(* IEC 61131-3 sources: plc-st-coding-agent/progress/evidence/f14_v3_parallel_20261112/jobs/codex_minimax-m27, 122 files *)

(* ---- public-easy-01.candidate_01.st ---- *)
FUNCTION_BLOCK FillingLineControl
VAR
    currentState : INT := 0;
END_VAR

CASE currentState OF
    0:
        Pump_Motor := FALSE;
        Filling_Valve := FALSE;
        Capping_Machine := FALSE;
        Packing_Machine := FALSE;
        Completion_Light := FALSE;

        IF bottleSensor THEN
            currentState := 1;
        END_IF;

    1:
        Pump_Motor := TRUE;

        IF cleaningConfirmButton THEN
            currentState := 2;
        END_IF;

    2:
        Pump_Motor := FALSE;
        Filling_Valve := TRUE;

        IF fillingConfirmButton THEN
            currentState := 3;
        END_IF;

    3:
        Filling_Valve := FALSE;
        Capping_Machine := TRUE;

        IF cappingConfirmButton THEN
            currentState := 4;
        END_IF;

    4:
        Capping_Machine := FALSE;
        Packing_Machine := TRUE;

        IF packingConfirmButton THEN
            currentState := 5;
        END_IF;

    5:
        Packing_Machine := FALSE;
        Completion_Light := TRUE;

        IF finishedButton THEN
            currentState := 0;
        END_IF;
END_CASE;
END_FUNCTION_BLOCK

(* ---- public-easy-01.candidate_02.st ---- *)
FUNCTION_BLOCK FillingLineControl
VAR_INPUT
    bottleSensor : BOOL;
    cleaningConfirmButton : BOOL;
    fillingConfirmButton : BOOL;
    cappingConfirmButton : BOOL;
    packingConfirmButton : BOOL;
    finishedButton : BOOL;
END_VAR
VAR_OUTPUT
    Pump_Motor : BOOL;
    Filling_Valve : BOOL;
    Capping_Machine : BOOL;
    Packing_Machine : BOOL;
    Completion_Light : BOOL;
END_VAR
VAR
    currentState : INT := 0;
END_VAR

CASE currentState OF
    0:
        Pump_Motor := FALSE;
        Filling_Valve := FALSE;
        Capping_Machine := FALSE;
        Packing_Machine := FALSE;
        Completion_Light := FALSE;

        IF bottleSensor THEN
            currentState := 1;
        END_IF;

    1:
        Pump_Motor := TRUE;

        IF cleaningConfirmButton THEN
            currentState := 2;
        END_IF;

    2:
        Pump_Motor := FALSE;
        Filling_Valve := TRUE;

        IF fillingConfirmButton THEN
            currentState := 3;
        END_IF;

    3:
        Filling_Valve := FALSE;
        Capping_Machine := TRUE;

        IF cappingConfirmButton THEN
            currentState := 4;
        END_IF;

    4:
        Capping_Machine := FALSE;
        Packing_Machine := TRUE;

        IF packingConfirmButton THEN
            currentState := 5;
        END_IF;

    5:
        Packing_Machine := FALSE;
        Completion_Light := TRUE;

        IF finishedButton THEN
            currentState := 0;
        END_IF;
END_CASE;
END_FUNCTION_BLOCK

(* ---- public-easy-01.raw_candidate_01.st ---- *)
FUNCTION_BLOCK FillingLineControl
VAR
    currentState : INT := 0;
END_VAR

CASE currentState OF
    0:
        Pump_Motor := FALSE;
        Filling_Valve := FALSE;
        Capping_Machine := FALSE;
        Packing_Machine := FALSE;
        Completion_Light := FALSE;

        IF bottleSensor THEN
            currentState := 1;
        END_IF;

    1:
        Pump_Motor := TRUE;

        IF cleaningConfirmButton THEN
            currentState := 2;
        END_IF;

    2:
        Pump_Motor := FALSE;
        Filling_Valve := TRUE;

        IF fillingConfirmButton THEN
            currentState := 3;
        END_IF;

    3:
        Filling_Valve := FALSE;
        Capping_Machine := TRUE;

        IF cappingConfirmButton THEN
            currentState := 4;
        END_IF;

    4:
        Capping_Machine := FALSE;
        Packing_Machine := TRUE;

        IF packingConfirmButton THEN
            currentState := 5;
        END_IF;

    5:
        Packing_Machine := FALSE;
        Completion_Light := TRUE;

        IF finishedButton THEN
            currentState := 0;
        END_IF;
END_CASE;
END_FUNCTION_BLOCK

(* ---- public-easy-01.raw_candidate_02.st ---- *)
FUNCTION_BLOCK FillingLineControl
VAR_INPUT
    bottleSensor : BOOL;
    cleaningConfirmButton : BOOL;
    fillingConfirmButton : BOOL;
    cappingConfirmButton : BOOL;
    packingConfirmButton : BOOL;
    finishedButton : BOOL;
END_VAR
VAR_OUTPUT
    Pump_Motor : BOOL;
    Filling_Valve : BOOL;
    Capping_Machine : BOOL;
    Packing_Machine : BOOL;
    Completion_Light : BOOL;
END_VAR
VAR
    currentState : INT := 0;
END_VAR

CASE currentState OF
    0:
        Pump_Motor := FALSE;
        Filling_Valve := FALSE;
        Capping_Machine := FALSE;
        Packing_Machine := FALSE;
        Completion_Light := FALSE;

        IF bottleSensor THEN
            currentState := 1;
        END_IF;

    1:
        Pump_Motor := TRUE;

        IF cleaningConfirmButton THEN
            currentState := 2;
        END_IF;

    2:
        Pump_Motor := FALSE;
        Filling_Valve := TRUE;

        IF fillingConfirmButton THEN
            currentState := 3;
        END_IF;

    3:
        Filling_Valve := FALSE;
        Capping_Machine := TRUE;

        IF cappingConfirmButton THEN
            currentState := 4;
        END_IF;

    4:
        Capping_Machine := FALSE;
        Packing_Machine := TRUE;

        IF packingConfirmButton THEN
            currentState := 5;
        END_IF;

    5:
        Packing_Machine := FALSE;
        Completion_Light := TRUE;

        IF finishedButton THEN
            currentState := 0;
        END_IF;
END_CASE;
END_FUNCTION_BLOCK

(* ---- public-easy-02.candidate_01.st ---- *)
FUNCTION_BLOCK FB_DualWordEdgeDetection
VAR_INPUT
END_VAR

VAR_OUTPUT
    hasChanged       : BOOL  := FALSE;
    hasRisingEdges   : BOOL  := FALSE;
    risingBits       : DWORD := 0;
    noOfRisingBits   : USINT := 0;
    hasFallingEdges  : BOOL  := FALSE;
    fallingBits      : DWORD := 0;
    noOfFallingBits  : USINT := 0;
END_VAR

VAR
    prevValue : DWORD := 0;
    bitMask   : DWORD;
    bitCount  : USINT;
END_VAR

// Detect rising edges: current=1 AND previous=0
risingBits := value AND (NOT prevValue);

// Detect falling edges: current=0 AND previous=1
fallingBits := (NOT value) AND prevValue;

// Set change indicators
hasChanged := (risingBits OR fallingBits) <> 0;
hasRisingEdges := risingBits <> 0;
hasFallingEdges := fallingBits <> 0;

// Count rising bits
bitMask := risingBits;
noOfRisingBits := 0;
FOR bitCount := 0 TO 31 DO
    IF (bitMask AND 1) = 1 THEN
        noOfRisingBits := noOfRisingBits + 1;
    END_IF;
    bitMask := SHR(bitMask, 1);
END_FOR;

// Count falling bits
bitMask := fallingBits;
noOfFallingBits := 0;
FOR bitCount := 0 TO 31 DO
    IF (bitMask AND 1) = 1 THEN
        noOfFallingBits := noOfFallingBits + 1;
    END_IF;
    bitMask := SHR(bitMask, 1);
END_FOR;

// Store current value for next scan
prevValue := value;

END_FUNCTION_BLOCK

(* ---- public-easy-02.candidate_02.st ---- *)
FUNCTION_BLOCK FB_DualWordEdgeDetection
VAR_INPUT
    value : DWORD;
END_VAR

VAR_OUTPUT
    hasChanged       : BOOL  := FALSE;
    hasRisingEdges   : BOOL  := FALSE;
    risingBits       : DWORD := 0;
    noOfRisingBits   : USINT := 0;
    hasFallingEdges  : BOOL  := FALSE;
    fallingBits      : DWORD := 0;
    noOfFallingBits  : USINT := 0;
END_VAR

VAR
    prevValue : DWORD := 0;
    tmpBits   : DWORD;
END_VAR

risingBits := value AND (NOT prevValue);
fallingBits := (NOT value) AND prevValue;

hasChanged := risingBits <> 0 OR fallingBits <> 0;
hasRisingEdges := risingBits <> 0;
hasFallingEdges := fallingBits <> 0;

tmpBits := risingBits;
noOfRisingBits := 0;
WHILE tmpBits <> 0 DO
    noOfRisingBits := noOfRisingBits + 1;
    tmpBits := SHR(tmpBits, 1);
END_WHILE;

tmpBits := fallingBits;
noOfFallingBits := 0;
WHILE tmpBits <> 0 DO
    noOfFallingBits := noOfFallingBits + 1;
    tmpBits := SHR(tmpBits, 1);
END_WHILE;

prevValue := value;

END_FUNCTION_BLOCK

(* ---- public-easy-02.raw_candidate_01.st ---- *)
FUNCTION_BLOCK FB_DualWordEdgeDetection
VAR_INPUT
END_VAR

VAR_OUTPUT
    hasChanged       : BOOL  := FALSE;
    hasRisingEdges   : BOOL  := FALSE;
    risingBits       : DWORD := 0;
    noOfRisingBits   : USINT := 0;
    hasFallingEdges  : BOOL  := FALSE;
    fallingBits      : DWORD := 0;
    noOfFallingBits  : USINT := 0;
END_VAR

VAR
    prevValue : DWORD := 0;
    bitMask   : DWORD;
    bitCount  : USINT;
END_VAR

// Detect rising edges: current=1 AND previous=0
risingBits := value AND (NOT prevValue);

// Detect falling edges: current=0 AND previous=1
fallingBits := (NOT value) AND prevValue;

// Set change indicators
hasChanged := (risingBits OR fallingBits) <> 0;
hasRisingEdges := risingBits <> 0;
hasFallingEdges := fallingBits <> 0;

// Count rising bits
bitMask := risingBits;
noOfRisingBits := 0;
FOR bitCount := 0 TO 31 DO
    IF (bitMask AND 1) = 1 THEN
        noOfRisingBits := noOfRisingBits + 1;
    END_IF;
    bitMask := SHR(bitMask, 1);
END_FOR;

// Count falling bits
bitMask := fallingBits;
noOfFallingBits := 0;
FOR bitCount := 0 TO 31 DO
    IF (bitMask AND 1) = 1 THEN
        noOfFallingBits := noOfFallingBits + 1;
    END_IF;
    bitMask := SHR(bitMask, 1);
END_FOR;

// Store current value for next scan
prevValue := value;

END_FUNCTION_BLOCK

(* ---- public-easy-02.raw_candidate_02.st ---- *)
FUNCTION_BLOCK FB_DualWordEdgeDetection
VAR_INPUT
    value : DWORD;
END_VAR

VAR_OUTPUT
    hasChanged       : BOOL  := FALSE;
    hasRisingEdges   : BOOL  := FALSE;
    risingBits       : DWORD := 0;
    noOfRisingBits   : USINT := 0;
    hasFallingEdges  : BOOL  := FALSE;
    fallingBits      : DWORD := 0;
    noOfFallingBits  : USINT := 0;
END_VAR

VAR
    prevValue : DWORD := 0;
    tmpBits   : DWORD;
END_VAR

risingBits := value AND (NOT prevValue);
fallingBits := (NOT value) AND prevValue;

hasChanged := risingBits <> 0 OR fallingBits <> 0;
hasRisingEdges := risingBits <> 0;
hasFallingEdges := fallingBits <> 0;

tmpBits := risingBits;
noOfRisingBits := 0;
WHILE tmpBits <> 0 DO
    noOfRisingBits := noOfRisingBits + 1;
    tmpBits := SHR(tmpBits, 1);
END_WHILE;

tmpBits := fallingBits;
noOfFallingBits := 0;
WHILE tmpBits <> 0 DO
    noOfFallingBits := noOfFallingBits + 1;
    tmpBits := SHR(tmpBits, 1);
END_WHILE;

prevValue := value;

END_FUNCTION_BLOCK

(* ---- public-easy-04.candidate_01.st ---- *)
FUNCTION_BLOCK JamPumpControl
VAR_INPUT
    VISCOSITY_OK     : BOOL;
    PASTE_E_STOP_NC  : BOOL;
    DebounceTime     : TIME;
    CycleTime        : TIME;
END_VAR

VAR_OUTPUT
    VFD_RUN          : BOOL := FALSE;
    PUMP_MAINT_DUE   : BOOL := FALSE;
    PUMP_RUNTIME_ACC : LTIME := LTIME#0s;
END_VAR

VAR
    ViscosityValid        : BOOL := FALSE;
    ViscosityDebounceTmr  : LTIME := LTIME#0s;
END_VAR

// Viscosity debouncing
IF VISCOSITY_OK THEN
    IF NOT ViscosityValid THEN
        ViscosityDebounceTmr := ViscosityDebounceTmr + LTIME(CycleTime);
        IF ViscosityDebounceTmr >= LTIME(DebounceTime) THEN
            ViscosityValid := TRUE;
            ViscosityDebounceTmr := LTIME#0s;
        END_IF;
    END_IF;
ELSE
    ViscosityValid := FALSE;
    ViscosityDebounceTmr := LTIME#0s;
END_IF;

// Safety permissive: E-stop AND valid viscosity
IF PASTE_E_STOP_NC AND ViscosityValid THEN
    VFD_RUN := TRUE;
ELSE
    VFD_RUN := FALSE;
END_IF;

// Runtime accumulation while running
IF VFD_RUN THEN
    PUMP_RUNTIME_ACC := PUMP_RUNTIME_ACC + LTIME(CycleTime);
END_IF;

// Maintenance due at 500 hours
PUMP_MAINT_DUE := (PUMP_RUNTIME_ACC >= LTIME#500h);

END_FUNCTION_BLOCK

(* ---- public-easy-04.candidate_02.st ---- *)
FUNCTION_BLOCK JamPumpControl
VAR_INPUT
    VISCOSITY_OK    : BOOL;
    PASTE_E_STOP_NC : BOOL;
    DebounceTime    : TIME;
    CycleTime       : TIME;
END_VAR

VAR_OUTPUT
    VFD_RUN          : BOOL := FALSE;
    PUMP_MAINT_DUE   : BOOL := FALSE;
    PUMP_RUNTIME_ACC : LTIME := LTIME#0s;
END_VAR

VAR
    ViscosityValid       : BOOL := FALSE;
    ViscosityDebounceTmr : LTIME := LTIME#0s;
END_VAR

IF VISCOSITY_OK THEN
    IF NOT ViscosityValid THEN
        ViscosityDebounceTmr := ViscosityDebounceTmr + CycleTime;
        IF ViscosityDebounceTmr >= DebounceTime THEN
            ViscosityValid := TRUE;
            ViscosityDebounceTmr := LTIME#0s;
        END_IF;
    END_IF;
ELSE
    ViscosityValid := FALSE;
    ViscosityDebounceTmr := LTIME#0s;
END_IF;

IF PASTE_E_STOP_NC AND ViscosityValid THEN
    VFD_RUN := TRUE;
ELSE
    VFD_RUN := FALSE;
END_IF;

IF VFD_RUN THEN
    PUMP_RUNTIME_ACC := PUMP_RUNTIME_ACC + CycleTime;
END_IF;

PUMP_MAINT_DUE := (PUMP_RUNTIME_ACC >= LTIME#500h);

END_FUNCTION_BLOCK

(* ---- public-easy-04.raw_candidate_01.st ---- *)
FUNCTION_BLOCK JamPumpControl
VAR_INPUT
    VISCOSITY_OK     : BOOL;
    PASTE_E_STOP_NC  : BOOL;
    DebounceTime     : TIME;
    CycleTime        : TIME;
END_VAR

VAR_OUTPUT
    VFD_RUN          : BOOL := FALSE;
    PUMP_MAINT_DUE   : BOOL := FALSE;
    PUMP_RUNTIME_ACC : LTIME := LTIME#0s;
END_VAR

VAR
    ViscosityValid        : BOOL := FALSE;
    ViscosityDebounceTmr  : LTIME := LTIME#0s;
END_VAR

// Viscosity debouncing
IF VISCOSITY_OK THEN
    IF NOT ViscosityValid THEN
        ViscosityDebounceTmr := ViscosityDebounceTmr + LTIME(CycleTime);
        IF ViscosityDebounceTmr >= LTIME(DebounceTime) THEN
            ViscosityValid := TRUE;
            ViscosityDebounceTmr := LTIME#0s;
        END_IF;
    END_IF;
ELSE
    ViscosityValid := FALSE;
    ViscosityDebounceTmr := LTIME#0s;
END_IF;

// Safety permissive: E-stop AND valid viscosity
IF PASTE_E_STOP_NC AND ViscosityValid THEN
    VFD_RUN := TRUE;
ELSE
    VFD_RUN := FALSE;
END_IF;

// Runtime accumulation while running
IF VFD_RUN THEN
    PUMP_RUNTIME_ACC := PUMP_RUNTIME_ACC + LTIME(CycleTime);
END_IF;

// Maintenance due at 500 hours
PUMP_MAINT_DUE := (PUMP_RUNTIME_ACC >= LTIME#500h);

END_FUNCTION_BLOCK

(* ---- public-easy-04.raw_candidate_02.st ---- *)
FUNCTION_BLOCK JamPumpControl
VAR_INPUT
    VISCOSITY_OK    : BOOL;
    PASTE_E_STOP_NC : BOOL;
    DebounceTime    : TIME;
    CycleTime       : TIME;
END_VAR

VAR_OUTPUT
    VFD_RUN          : BOOL := FALSE;
    PUMP_MAINT_DUE   : BOOL := FALSE;
    PUMP_RUNTIME_ACC : LTIME := LTIME#0s;
END_VAR

VAR
    ViscosityValid       : BOOL := FALSE;
    ViscosityDebounceTmr : LTIME := LTIME#0s;
END_VAR

IF VISCOSITY_OK THEN
    IF NOT ViscosityValid THEN
        ViscosityDebounceTmr := ViscosityDebounceTmr + CycleTime;
        IF ViscosityDebounceTmr >= DebounceTime THEN
            ViscosityValid := TRUE;
            ViscosityDebounceTmr := LTIME#0s;
        END_IF;
    END_IF;
ELSE
    ViscosityValid := FALSE;
    ViscosityDebounceTmr := LTIME#0s;
END_IF;

IF PASTE_E_STOP_NC AND ViscosityValid THEN
    VFD_RUN := TRUE;
ELSE
    VFD_RUN := FALSE;
END_IF;

IF VFD_RUN THEN
    PUMP_RUNTIME_ACC := PUMP_RUNTIME_ACC + CycleTime;
END_IF;

PUMP_MAINT_DUE := (PUMP_RUNTIME_ACC >= LTIME#500h);

END_FUNCTION_BLOCK

(* ---- public-easy-05.candidate_01.st ---- *)
FUNCTION_BLOCK WeldGapAlarm
VAR_INPUT
    Gap_Exceeded : BOOL;
    Weld_E_Stop_NC : BOOL;
    DebounceTime : TIME;
END_VAR

VAR_OUTPUT
    Operator_Alert : BOOL := FALSE;
    Weld_Soft_Start_Active : BOOL := TRUE;
END_VAR

VAR
    initTimer : TON;
    debounceTimer : TON;
    monitoringActive : BOOL := FALSE;
END_VAR

// E-Stop takes priority over all states
IF NOT Weld_E_Stop_NC THEN
    Operator_Alert := FALSE;
    Weld_Soft_Start_Active := FALSE;
    monitoringActive := FALSE;

    // Reset timers when E-Stop is active
    initTimer(IN := FALSE);
    debounceTimer(IN := FALSE);
    initTimer();
    debounceTimer();
    RETURN;
END_IF;

// Initialization phase: 5-second power-up inhibition
IF NOT monitoringActive THEN
    initTimer(IN := TRUE, PT := T#5S);
    initTimer();

    Operator_Alert := FALSE;
    Weld_Soft_Start_Active := TRUE;

    IF initTimer.Q THEN
        monitoringActive := TRUE;
        Weld_Soft_Start_Active := FALSE;

        // Reset timers upon entering monitoring
        initTimer(IN := FALSE);
        debounceTimer(IN := FALSE);
        initTimer();
        debounceTimer();
    END_IF;

    initTimer(IN := FALSE);
    initTimer();
    RETURN;
END_IF;

// Normal gap monitoring with debounce
IF NOT Gap_Exceeded THEN
    Operator_Alert := FALSE;
    debounceTimer(IN := FALSE);
    debounceTimer();
ELSE
    debounceTimer(IN := TRUE, PT := DebounceTime);
    debounceTimer();

    IF debounceTimer.Q THEN
        Operator_Alert := TRUE;
    END_IF;
END_IF;

END_FUNCTION_BLOCK

(* ---- public-easy-05.candidate_02.st ---- *)
FUNCTION_BLOCK WeldGapAlarm
VAR_INPUT
    Gap_Exceeded : BOOL;
    Weld_E_Stop_NC : BOOL;
    DebounceTime : TIME;
END_VAR

VAR_OUTPUT
    Operator_Alert : BOOL := FALSE;
    Weld_Soft_Start_Active : BOOL := TRUE;
END_VAR

VAR
    initTimer : TON;
    debounceTimer : TON;
    state : UINT := 0;
END_VAR

IF NOT Weld_E_Stop_NC THEN
    Operator_Alert := FALSE;
    Weld_Soft_Start_Active := FALSE;
    state := 0;
    initTimer(IN := FALSE);
    debounceTimer(IN := FALSE);
    initTimer();
    debounceTimer();
    RETURN;
END_IF;

IF state = 0 THEN
    initTimer(IN := TRUE, PT := T#5S);
    initTimer();
    Operator_Alert := FALSE;
    Weld_Soft_Start_Active := TRUE;

    IF initTimer.Q THEN
        state := 1;
        initTimer(IN := FALSE);
        debounceTimer(IN := FALSE);
        initTimer();
        debounceTimer();
    END_IF;
    RETURN;
END_IF;

IF state = 1 THEN
    Weld_Soft_Start_Active := FALSE;

    IF NOT Gap_Exceeded THEN
        Operator_Alert := FALSE;
        debounceTimer(IN := FALSE);
        debounceTimer();
    ELSE
        debounceTimer(IN := TRUE, PT := DebounceTime);
        debounceTimer();

        IF debounceTimer.Q THEN
            Operator_Alert := TRUE;
        END_IF;
    END_IF;
END_IF;

END_FUNCTION_BLOCK

(* ---- public-easy-05.raw_candidate_01.st ---- *)
FUNCTION_BLOCK WeldGapAlarm
VAR_INPUT
    Gap_Exceeded : BOOL;
    Weld_E_Stop_NC : BOOL;
    DebounceTime : TIME;
END_VAR

VAR_OUTPUT
    Operator_Alert : BOOL := FALSE;
    Weld_Soft_Start_Active : BOOL := TRUE;
END_VAR

VAR
    initTimer : TON;
    debounceTimer : TON;
    monitoringActive : BOOL := FALSE;
END_VAR

// E-Stop takes priority over all states
IF NOT Weld_E_Stop_NC THEN
    Operator_Alert := FALSE;
    Weld_Soft_Start_Active := FALSE;
    monitoringActive := FALSE;

    // Reset timers when E-Stop is active
    initTimer(IN := FALSE);
    debounceTimer(IN := FALSE);
    initTimer();
    debounceTimer();
    RETURN;
END_IF;

// Initialization phase: 5-second power-up inhibition
IF NOT monitoringActive THEN
    initTimer(IN := TRUE, PT := T#5S);
    initTimer();

    Operator_Alert := FALSE;
    Weld_Soft_Start_Active := TRUE;

    IF initTimer.Q THEN
        monitoringActive := TRUE;
        Weld_Soft_Start_Active := FALSE;

        // Reset timers upon entering monitoring
        initTimer(IN := FALSE);
        debounceTimer(IN := FALSE);
        initTimer();
        debounceTimer();
    END_IF;

    initTimer(IN := FALSE);
    initTimer();
    RETURN;
END_IF;

// Normal gap monitoring with debounce
IF NOT Gap_Exceeded THEN
    Operator_Alert := FALSE;
    debounceTimer(IN := FALSE);
    debounceTimer();
ELSE
    debounceTimer(IN := TRUE, PT := DebounceTime);
    debounceTimer();

    IF debounceTimer.Q THEN
        Operator_Alert := TRUE;
    END_IF;
END_IF;

END_FUNCTION_BLOCK

(* ---- public-easy-05.raw_candidate_02.st ---- *)
FUNCTION_BLOCK WeldGapAlarm
VAR_INPUT
    Gap_Exceeded : BOOL;
    Weld_E_Stop_NC : BOOL;
    DebounceTime : TIME;
END_VAR

VAR_OUTPUT
    Operator_Alert : BOOL := FALSE;
    Weld_Soft_Start_Active : BOOL := TRUE;
END_VAR

VAR
    initTimer : TON;
    debounceTimer : TON;
    state : UINT := 0;
END_VAR

IF NOT Weld_E_Stop_NC THEN
    Operator_Alert := FALSE;
    Weld_Soft_Start_Active := FALSE;
    state := 0;
    initTimer(IN := FALSE);
    debounceTimer(IN := FALSE);
    initTimer();
    debounceTimer();
    RETURN;
END_IF;

IF state = 0 THEN
    initTimer(IN := TRUE, PT := T#5S);
    initTimer();
    Operator_Alert := FALSE;
    Weld_Soft_Start_Active := TRUE;

    IF initTimer.Q THEN
        state := 1;
        initTimer(IN := FALSE);
        debounceTimer(IN := FALSE);
        initTimer();
        debounceTimer();
    END_IF;
    RETURN;
END_IF;

IF state = 1 THEN
    Weld_Soft_Start_Active := FALSE;

    IF NOT Gap_Exceeded THEN
        Operator_Alert := FALSE;
        debounceTimer(IN := FALSE);
        debounceTimer();
    ELSE
        debounceTimer(IN := TRUE, PT := DebounceTime);
        debounceTimer();

        IF debounceTimer.Q THEN
            Operator_Alert := TRUE;
        END_IF;
    END_IF;
END_IF;

END_FUNCTION_BLOCK

(* ---- public-easy-06.candidate_01.st ---- *)
FUNCTION_BLOCK AerationBlowerControl
VAR_INPUT
    DO_LOW : BOOL;
    AERATION_E_STOP_NC : BOOL;
END_VAR

VAR_OUTPUT
    BLOWER_RUN : BOOL := FALSE;
    AERATION_BLOWER_CYCLE_COUNT : UINT := 0;
END_VAR

VAR
    StartTimer : TON;
    WasRunning : BOOL := FALSE;
END_VAR

    StartTimer(IN := DO_LOW AND AERATION_E_STOP_NC, PT := T#5S);

    BLOWER_RUN := StartTimer.Q;

    IF BLOWER_RUN AND NOT WasRunning THEN
        AERATION_BLOWER_CYCLE_COUNT := AERATION_BLOWER_CYCLE_COUNT + 1;
    END_IF;

    WasRunning := BLOWER_RUN;
END_FUNCTION_BLOCK

(* ---- public-easy-06.raw_candidate_01.st ---- *)
FUNCTION_BLOCK AerationBlowerControl
VAR_INPUT
    DO_LOW : BOOL;
    AERATION_E_STOP_NC : BOOL;
END_VAR

VAR_OUTPUT
    BLOWER_RUN : BOOL := FALSE;
    AERATION_BLOWER_CYCLE_COUNT : UINT := 0;
END_VAR

VAR
    StartTimer : TON;
    WasRunning : BOOL := FALSE;
END_VAR

    StartTimer(IN := DO_LOW AND AERATION_E_STOP_NC, PT := T#5S);

    BLOWER_RUN := StartTimer.Q;

    IF BLOWER_RUN AND NOT WasRunning THEN
        AERATION_BLOWER_CYCLE_COUNT := AERATION_BLOWER_CYCLE_COUNT + 1;
    END_IF;

    WasRunning := BLOWER_RUN;
END_FUNCTION_BLOCK

(* ---- public-hard-01.candidate_01.st ---- *)
FUNCTION_BLOCK MaterialProportioningControl
VAR_INPUT
    estop           : BOOL;
    opeMode         : BOOL;
    valveAStart     : BOOL;
    valveBStart     : BOOL;
    valveCStart     : BOOL;
    valveDStart     : BOOL;
    mixMotorStart   : BOOL;
    autoStart       : BOOL;
    processMode     : BOOL;
    levelSensor     : INT;
    mixMotorComplete: BOOL;
END_VAR

VAR_OUTPUT
    valveARun       : BOOL;
    valveBRun       : BOOL;
    valveCRun       : BOOL;
    valveDRun       : BOOL;
    mixMotorRun     : BOOL;
END_VAR

VAR
    prevValveAStart     : BOOL := FALSE;
    prevValveBStart     : BOOL := FALSE;
    prevValveCStart     : BOOL := FALSE;
    prevValveDStart     : BOOL := FALSE;
    prevMixMotorStart   : BOOL := FALSE;
    prevAutoStart       : BOOL := FALSE;
    autoState           : INT := 0;
    autoRunning         : BOOL := FALSE;
END_VAR

// Emergency Stop - stops all equipment immediately
IF NOT estop THEN
    valveARun   := FALSE;
    valveBRun   := FALSE;
    valveCRun   := FALSE;
    valveDRun   := FALSE;
    mixMotorRun := FALSE;
    autoRunning := FALSE;
    autoState   := 0;
    RETURN;
END_IF;

// Manual Mode
IF NOT opeMode THEN
    // Rising edge detection for Valve A toggle
    IF valveAStart AND NOT prevValveAStart THEN
        valveARun := NOT valveARun;
    END_IF;
    prevValveAStart := valveAStart;

    // Rising edge detection for Valve B toggle
    IF valveBStart AND NOT prevValveBStart THEN
        valveBRun := NOT valveBRun;
    END_IF;
    prevValveBStart := valveBStart;

    // Rising edge detection for Valve C toggle
    IF valveCStart AND NOT prevValveCStart THEN
        valveCRun := NOT valveCRun;
    END_IF;
    prevValveCStart := valveCStart;

    // Rising edge detection for Valve D toggle
    IF valveDStart AND NOT prevValveDStart THEN
        valveDRun := NOT valveDRun;
    END_IF;
    prevValveDStart := valveDStart;

    // Rising edge detection for Mixing Motor toggle
    IF mixMotorStart AND NOT prevMixMotorStart THEN
        mixMotorRun := NOT mixMotorRun;
    END_IF;
    prevMixMotorStart := mixMotorStart;

// Automatic Mode
ELSE
    // Rising edge detection for autoStart
    IF autoStart AND NOT prevAutoStart AND NOT autoRunning THEN
        autoRunning := TRUE;
        autoState   := 1;
    END_IF;
    prevAutoStart := autoStart;

    // State machine for automatic process flow
    IF autoRunning THEN
        CASE autoState OF
            1: // Open Valve A
                valveARun := TRUE;
                IF levelSensor >= 50 THEN
                    valveARun := FALSE;
                    autoState := 2;
                END_IF;

            2: // Open Valve B, wait for level 80cm
                valveBRun := TRUE;
                IF levelSensor >= 80 THEN
                    valveBRun := FALSE;
                    IF processMode THEN
                        autoState := 3;
                    ELSE
                        autoState := 4;
                    END_IF;
                END_IF;

            3: // Open Valve C (processMode=true), wait for level 100cm
                valveCRun := TRUE;
                IF levelSensor >= 100 THEN
                    valveCRun := FALSE;
                    autoState := 4;
                END_IF;

            4: // Start mixing motor
                mixMotorRun := TRUE;
                IF mixMotorComplete THEN
                    mixMotorRun := FALSE;
                    autoState := 5;
                END_IF;

            5: // Open Valve D, end automatic process
                valveDRun  := TRUE;
                autoRunning := FALSE;
                autoState   := 0;
        END_CASE;
    END_IF;
END_IF;

END_FUNCTION_BLOCK

(* ---- public-hard-01.candidate_02.st ---- *)
FUNCTION_BLOCK MaterialProportioningControl
VAR_INPUT
    estop           : BOOL;
    opeMode         : BOOL;
    valveAStart     : BOOL;
    valveBStart     : BOOL;
    valveCStart     : BOOL;
    valveDStart     : BOOL;
    mixMotorStart   : BOOL;
    autoStart       : BOOL;
    processMode     : BOOL;
    levelSensor     : INT;
    mixMotorComplete: BOOL;
END_VAR

VAR_OUTPUT
    valveARun       : BOOL;
    valveBRun       : BOOL;
    valveCRun       : BOOL;
    valveDRun       : BOOL;
    mixMotorRun     : BOOL;
END_VAR

VAR
    prevValveAStart     : BOOL := FALSE;
    prevValveBStart     : BOOL := FALSE;
    prevValveCStart     : BOOL := FALSE;
    prevValveDStart     : BOOL := FALSE;
    prevMixMotorStart   : BOOL := FALSE;
    prevAutoStart       : BOOL := FALSE;
    autoState           : INT := 0;
END_VAR

// Emergency Stop - stops all equipment immediately, but preserve autoState for resumption
IF NOT estop THEN
    valveARun   := FALSE;
    valveBRun   := FALSE;
    valveCRun   := FALSE;
    valveDRun   := FALSE;
    mixMotorRun := FALSE;
    RETURN;
END_IF;

// Manual Mode
IF NOT opeMode THEN
    // Rising edge detection for Valve A toggle
    IF valveAStart AND NOT prevValveAStart THEN
        valveARun := NOT valveARun;
    END_IF;
    prevValveAStart := valveAStart;

    // Rising edge detection for Valve B toggle
    IF valveBStart AND NOT prevValveBStart THEN
        valveBRun := NOT valveBRun;
    END_IF;
    prevValveBStart := valveBStart;

    // Rising edge detection for Valve C toggle
    IF valveCStart AND NOT prevValveCStart THEN
        valveCRun := NOT valveCRun;
    END_IF;
    prevValveCStart := valveCStart;

    // Rising edge detection for Valve D toggle
    IF valveDStart AND NOT prevValveDStart THEN
        valveDRun := NOT valveDRun;
    END_IF;
    prevValveDStart := valveDStart;

    // Rising edge detection for Mixing Motor toggle
    IF mixMotorStart AND NOT prevMixMotorStart THEN
        mixMotorRun := NOT mixMotorRun;
    END_IF;
    prevMixMotorStart := mixMotorStart;

// Automatic Mode
ELSE
    // Rising edge detection for autoStart - initiates or resumes automatic process
    IF autoStart AND NOT prevAutoStart THEN
        IF autoState = 0 THEN
            autoState := 1;
        END_IF;
    END_IF;
    prevAutoStart := autoStart;

    // State machine for automatic process flow
    CASE autoState OF
        1: // Open Valve A, wait for level >= 50cm
            valveARun := TRUE;
            valveBRun := FALSE;
            valveCRun := FALSE;
            valveDRun := FALSE;
            mixMotorRun := FALSE;
            IF levelSensor >= 50 THEN
                valveARun := FALSE;
                autoState := 2;
            END_IF;

        2: // Open Valve B, wait for level >= 80cm
            valveARun := FALSE;
            valveBRun := TRUE;
            valveCRun := FALSE;
            valveDRun := FALSE;
            mixMotorRun := FALSE;
            IF levelSensor >= 80 THEN
                valveBRun := FALSE;
                IF processMode THEN
                    autoState := 3;
                ELSE
                    autoState := 4;
                END_IF;
            END_IF;

        3: // Open Valve C (processMode=true), wait for level >= 100cm
            valveARun := FALSE;
            valveBRun := FALSE;
            valveCRun := TRUE;
            valveDRun := FALSE;
            mixMotorRun := FALSE;
            IF levelSensor >= 100 THEN
                valveCRun := FALSE;
                autoState := 4;
            END_IF;

        4: // Start mixing motor, wait for mixMotorComplete
            valveARun := FALSE;
            valveBRun := FALSE;
            valveCRun := FALSE;
            valveDRun := FALSE;
            mixMotorRun := TRUE;
            IF mixMotorComplete THEN
                mixMotorRun := FALSE;
                autoState := 5;
            END_IF;

        5: // Open Valve D, end automatic process
            valveARun := FALSE;
            valveBRun := FALSE;
            valveCRun := FALSE;
            valveDRun := TRUE;
            mixMotorRun := FALSE;
            autoState := 0;
    END_CASE;
END_IF;

END_FUNCTION_BLOCK

(* ---- public-hard-01.raw_candidate_01.st ---- *)
FUNCTION_BLOCK MaterialProportioningControl
VAR_INPUT
    estop           : BOOL;
    opeMode         : BOOL;
    valveAStart     : BOOL;
    valveBStart     : BOOL;
    valveCStart     : BOOL;
    valveDStart     : BOOL;
    mixMotorStart   : BOOL;
    autoStart       : BOOL;
    processMode     : BOOL;
    levelSensor     : INT;
    mixMotorComplete: BOOL;
END_VAR

VAR_OUTPUT
    valveARun       : BOOL;
    valveBRun       : BOOL;
    valveCRun       : BOOL;
    valveDRun       : BOOL;
    mixMotorRun     : BOOL;
END_VAR

VAR
    prevValveAStart     : BOOL := FALSE;
    prevValveBStart     : BOOL := FALSE;
    prevValveCStart     : BOOL := FALSE;
    prevValveDStart     : BOOL := FALSE;
    prevMixMotorStart   : BOOL := FALSE;
    prevAutoStart       : BOOL := FALSE;
    autoState           : INT := 0;
    autoRunning         : BOOL := FALSE;
END_VAR

// Emergency Stop - stops all equipment immediately
IF NOT estop THEN
    valveARun   := FALSE;
    valveBRun   := FALSE;
    valveCRun   := FALSE;
    valveDRun   := FALSE;
    mixMotorRun := FALSE;
    autoRunning := FALSE;
    autoState   := 0;
    RETURN;
END_IF

// Manual Mode
IF NOT opeMode THEN
    // Rising edge detection for Valve A toggle
    IF valveAStart AND NOT prevValveAStart THEN
        valveARun := NOT valveARun;
    END_IF;
    prevValveAStart := valveAStart;

    // Rising edge detection for Valve B toggle
    IF valveBStart AND NOT prevValveBStart THEN
        valveBRun := NOT valveBRun;
    END_IF;
    prevValveBStart := valveBStart;

    // Rising edge detection for Valve C toggle
    IF valveCStart AND NOT prevValveCStart THEN
        valveCRun := NOT valveCRun;
    END_IF;
    prevValveCStart := valveCStart;

    // Rising edge detection for Valve D toggle
    IF valveDStart AND NOT prevValveDStart THEN
        valveDRun := NOT valveDRun;
    END_IF;
    prevValveDStart := valveDStart;

    // Rising edge detection for Mixing Motor toggle
    IF mixMotorStart AND NOT prevMixMotorStart THEN
        mixMotorRun := NOT mixMotorRun;
    END_IF;
    prevMixMotorStart := mixMotorStart;

// Automatic Mode
ELSE
    // Rising edge detection for autoStart
    IF autoStart AND NOT prevAutoStart AND NOT autoRunning THEN
        autoRunning := TRUE;
        autoState   := 1;
    END_IF;
    prevAutoStart := autoStart;

    // State machine for automatic process flow
    IF autoRunning THEN
        CASE autoState OF
            1: // Open Valve A
                valveARun := TRUE;
                IF levelSensor >= 50 THEN
                    valveARun := FALSE;
                    autoState := 2;
                END_IF;

            2: // Open Valve B, wait for level 80cm
                valveBRun := TRUE;
                IF levelSensor >= 80 THEN
                    valveBRun := FALSE;
                    IF processMode THEN
                        autoState := 3;
                    ELSE
                        autoState := 4;
                    END_IF;
                END_IF;

            3: // Open Valve C (processMode=true), wait for level 100cm
                valveCRun := TRUE;
                IF levelSensor >= 100 THEN
                    valveCRun := FALSE;
                    autoState := 4;
                END_IF;

            4: // Start mixing motor
                mixMotorRun := TRUE;
                IF mixMotorComplete THEN
                    mixMotorRun := FALSE;
                    autoState := 5;
                END_IF;

            5: // Open Valve D, end automatic process
                valveDRun  := TRUE;
                autoRunning := FALSE;
                autoState   := 0;
        END_CASE;
    END_IF;
END_IF;

END_FUNCTION_BLOCK

(* ---- public-hard-01.raw_candidate_02.st ---- *)
FUNCTION_BLOCK MaterialProportioningControl
VAR_INPUT
    estop           : BOOL;
    opeMode         : BOOL;
    valveAStart     : BOOL;
    valveBStart     : BOOL;
    valveCStart     : BOOL;
    valveDStart     : BOOL;
    mixMotorStart   : BOOL;
    autoStart       : BOOL;
    processMode     : BOOL;
    levelSensor     : INT;
    mixMotorComplete: BOOL;
END_VAR

VAR_OUTPUT
    valveARun       : BOOL;
    valveBRun       : BOOL;
    valveCRun       : BOOL;
    valveDRun       : BOOL;
    mixMotorRun     : BOOL;
END_VAR

VAR
    prevValveAStart     : BOOL := FALSE;
    prevValveBStart     : BOOL := FALSE;
    prevValveCStart     : BOOL := FALSE;
    prevValveDStart     : BOOL := FALSE;
    prevMixMotorStart   : BOOL := FALSE;
    prevAutoStart       : BOOL := FALSE;
    autoState           : INT := 0;
END_VAR

// Emergency Stop - stops all equipment immediately, but preserve autoState for resumption
IF NOT estop THEN
    valveARun   := FALSE;
    valveBRun   := FALSE;
    valveCRun   := FALSE;
    valveDRun   := FALSE;
    mixMotorRun := FALSE;
    RETURN;
END_IF;

// Manual Mode
IF NOT opeMode THEN
    // Rising edge detection for Valve A toggle
    IF valveAStart AND NOT prevValveAStart THEN
        valveARun := NOT valveARun;
    END_IF;
    prevValveAStart := valveAStart;

    // Rising edge detection for Valve B toggle
    IF valveBStart AND NOT prevValveBStart THEN
        valveBRun := NOT valveBRun;
    END_IF;
    prevValveBStart := valveBStart;

    // Rising edge detection for Valve C toggle
    IF valveCStart AND NOT prevValveCStart THEN
        valveCRun := NOT valveCRun;
    END_IF;
    prevValveCStart := valveCStart;

    // Rising edge detection for Valve D toggle
    IF valveDStart AND NOT prevValveDStart THEN
        valveDRun := NOT valveDRun;
    END_IF;
    prevValveDStart := valveDStart;

    // Rising edge detection for Mixing Motor toggle
    IF mixMotorStart AND NOT prevMixMotorStart THEN
        mixMotorRun := NOT mixMotorRun;
    END_IF;
    prevMixMotorStart := mixMotorStart;

// Automatic Mode
ELSE
    // Rising edge detection for autoStart - initiates or resumes automatic process
    IF autoStart AND NOT prevAutoStart THEN
        IF autoState = 0 THEN
            autoState := 1;
        END_IF;
    END_IF;
    prevAutoStart := autoStart;

    // State machine for automatic process flow
    CASE autoState OF
        1: // Open Valve A, wait for level >= 50cm
            valveARun := TRUE;
            valveBRun := FALSE;
            valveCRun := FALSE;
            valveDRun := FALSE;
            mixMotorRun := FALSE;
            IF levelSensor >= 50 THEN
                valveARun := FALSE;
                autoState := 2;
            END_IF;

        2: // Open Valve B, wait for level >= 80cm
            valveARun := FALSE;
            valveBRun := TRUE;
            valveCRun := FALSE;
            valveDRun := FALSE;
            mixMotorRun := FALSE;
            IF levelSensor >= 80 THEN
                valveBRun := FALSE;
                IF processMode THEN
                    autoState := 3;
                ELSE
                    autoState := 4;
                END_IF;
            END_IF;

        3: // Open Valve C (processMode=true), wait for level >= 100cm
            valveARun := FALSE;
            valveBRun := FALSE;
            valveCRun := TRUE;
            valveDRun := FALSE;
            mixMotorRun := FALSE;
            IF levelSensor >= 100 THEN
                valveCRun := FALSE;
                autoState := 4;
            END_IF;

        4: // Start mixing motor, wait for mixMotorComplete
            valveARun := FALSE;
            valveBRun := FALSE;
            valveCRun := FALSE;
            valveDRun := FALSE;
            mixMotorRun := TRUE;
            IF mixMotorComplete THEN
                mixMotorRun := FALSE;
                autoState := 5;
            END_IF;

        5: // Open Valve D, end automatic process
            valveARun := FALSE;
            valveBRun := FALSE;
            valveCRun := FALSE;
            valveDRun := TRUE;
            mixMotorRun := FALSE;
            autoState := 0;
    END_CASE;
END_IF;

END_FUNCTION_BLOCK

(* ---- public-hard-02.candidate_01.st ---- *)
FUNCTION_BLOCK FlexibleProcessingControl
VAR_INPUT
    processLength    : USINT;
    sensor1          : BOOL;
    sensor2          : BOOL;
    sensor3          : BOOL;
    sensor4          : BOOL;
    sensor5          : BOOL;
    station1Start    : BOOL;
    station2Complete : BOOL;
    station3Complete : BOOL;
    station4Complete : BOOL;
    processSequence  : ARRAY[1..8] OF USINT;
END_VAR
VAR_OUTPUT
    conveyorLeft  : BOOL;
    conveyorRight : BOOL;
END_VAR
VAR
    state            : INT;
    currentStation   : USINT;
    sequenceIndex    : USINT;
    targetStation    : USINT;
    prevSensor1      : BOOL;
    prevSensor2      : BOOL;
    prevSensor3      : BOOL;
    prevSensor4      : BOOL;
    prevSensor5      : BOOL;
    waitComplete     : BOOL;
END_VAR

(* State constants *)
CONSTANT
    IDLE          : INT := 0;
    LOADING       : INT := 1;
    MOVING        : INT := 2;
    WAIT_PROCESS  : INT := 3;
END_CONSTANT

(* Main logic *)
CASE state OF
    IDLE:
        conveyorLeft  := FALSE;
        conveyorRight := FALSE;
        IF sensor1 AND station1Start THEN
            sequenceIndex  := 1;
            targetStation := processSequence[1];
            currentStation := 1;
            state := LOADING;
        END_IF;

    LOADING:
        conveyorLeft  := FALSE;
        conveyorRight := FALSE;
        sequenceIndex := 1;
        targetStation := processSequence[1];
        currentStation := 1;
        state := MOVING;

    MOVING:
        (* Rising edge detection for sensors *)
        IF sensor1 AND NOT prevSensor1 THEN
            currentStation := 1;
        END_IF;
        IF sensor2 AND NOT prevSensor2 THEN
            currentStation := 2;
        END_IF;
        IF sensor3 AND NOT prevSensor3 THEN
            currentStation := 3;
        END_IF;
        IF sensor4 AND NOT prevSensor4 THEN
            currentStation := 4;
        END_IF;
        IF sensor5 AND NOT prevSensor5 THEN
            currentStation := 5;
        END_IF;

        (* Determine conveyor direction based on target vs current *)
        IF targetStation > currentStation THEN
            conveyorRight := TRUE;
            conveyorLeft  := FALSE;
        ELSIF targetStation < currentStation THEN
            conveyorLeft  := TRUE;
            conveyorRight := FALSE;
        ELSE
            conveyorLeft  := FALSE;
            conveyorRight := FALSE;
        END_IF;

        (* Check if product reached target station *)
        IF currentStation = targetStation THEN
            conveyorLeft  := FALSE;
            conveyorRight := FALSE;
            state := WAIT_PROCESS;
            waitComplete := FALSE;
        END_IF;

    WAIT_PROCESS:
        IF NOT waitComplete THEN
            waitComplete := TRUE;
        END_IF;

        IF waitComplete THEN
            IF targetStation = 2 AND station2Complete THEN
                sequenceIndex := sequenceIndex + 1;
                state := CHECK_SEQUENCE;
            ELSIF targetStation = 3 AND station3Complete THEN
                sequenceIndex := sequenceIndex + 1;
                state := CHECK_SEQUENCE;
            ELSIF targetStation = 4 AND station4Complete THEN
                sequenceIndex := sequenceIndex + 1;
                state := CHECK_SEQUENCE;
            ELSIF targetStation = 5 THEN
                sequenceIndex := sequenceIndex + 1;
                state := CHECK_SEQUENCE;
            END_IF;
        END_IF;

    CHECK_SEQUENCE:
        IF sequenceIndex > processLength THEN
            state := IDLE;
        ELSE
            targetStation := processSequence[sequenceIndex];
            state := MOVING;
        END_IF;
END_CASE;

(* Update previous sensor states *)
prevSensor1 := sensor1;
prevSensor2 := sensor2;
prevSensor3 := sensor3;
prevSensor4 := sensor4;
prevSensor5 := sensor5;

END_FUNCTION_BLOCK

(* ---- public-hard-02.candidate_02.st ---- *)
TYPE
    ProcessState : INT (
        IDLE          := 0,
        LOADING       := 1,
        MOVING        := 2,
        WAIT_PROCESS  := 3,
        CHECK_SEQUENCE:= 4
    );
END_TYPE;

FUNCTION_BLOCK FlexibleProcessingControl
VAR_INPUT
    processLength    : USINT;
    sensor1          : BOOL;
    sensor2          : BOOL;
    sensor3          : BOOL;
    sensor4          : BOOL;
    sensor5          : BOOL;
    station1Start    : BOOL;
    station2Complete : BOOL;
    station3Complete : BOOL;
    station4Complete : BOOL;
    processSequence  : ARRAY[1..8] OF USINT;
END_VAR
VAR_OUTPUT
    conveyorLeft  : BOOL;
    conveyorRight : BOOL;
END_VAR
VAR
    internalState     : ProcessState;
    currentStation    : USINT;
    sequenceIndex     : USINT;
    targetStation     : USINT;
    prevSensor1       : BOOL;
    prevSensor2       : BOOL;
    prevSensor3       : BOOL;
    prevSensor4       : BOOL;
    prevSensor5       : BOOL;
    waitComplete      : BOOL;
END_VAR

CASE internalState OF
    IDLE:
        conveyorLeft  := FALSE;
        conveyorRight := FALSE;
        IF sensor1 AND station1Start THEN
            sequenceIndex  := 1;
            targetStation := processSequence[1];
            currentStation := 1;
            internalState := LOADING;
        END_IF;

    LOADING:
        conveyorLeft  := FALSE;
        conveyorRight := FALSE;
        sequenceIndex := 1;
        targetStation := processSequence[1];
        currentStation := 1;
        internalState := MOVING;

    MOVING:
        IF sensor1 AND NOT prevSensor1 THEN
            currentStation := 1;
        END_IF;
        IF sensor2 AND NOT prevSensor2 THEN
            currentStation := 2;
        END_IF;
        IF sensor3 AND NOT prevSensor3 THEN
            currentStation := 3;
        END_IF;
        IF sensor4 AND NOT prevSensor4 THEN
            currentStation := 4;
        END_IF;
        IF sensor5 AND NOT prevSensor5 THEN
            currentStation := 5;
        END_IF;

        IF targetStation > currentStation THEN
            conveyorRight := TRUE;
            conveyorLeft  := FALSE;
        ELSIF targetStation < currentStation THEN
            conveyorLeft  := TRUE;
            conveyorRight := FALSE;
        ELSE
            conveyorLeft  := FALSE;
            conveyorRight := FALSE;
        END_IF;

        IF currentStation = targetStation THEN
            conveyorLeft  := FALSE;
            conveyorRight := FALSE;
            internalState := WAIT_PROCESS;
            waitComplete := FALSE;
        END_IF;

    WAIT_PROCESS:
        IF NOT waitComplete THEN
            waitComplete := TRUE;
        END_IF;

        IF waitComplete THEN
            IF targetStation = 2 AND station2Complete THEN
                sequenceIndex := sequenceIndex + 1;
                internalState := CHECK_SEQUENCE;
            ELSIF targetStation = 3 AND station3Complete THEN
                sequenceIndex := sequenceIndex + 1;
                internalState := CHECK_SEQUENCE;
            ELSIF targetStation = 4 AND station4Complete THEN
                sequenceIndex := sequenceIndex + 1;
                internalState := CHECK_SEQUENCE;
            ELSIF targetStation = 5 THEN
                sequenceIndex := sequenceIndex + 1;
                internalState := CHECK_SEQUENCE;
            END_IF;
        END_IF;

    CHECK_SEQUENCE:
        IF sequenceIndex > processLength THEN
            internalState := IDLE;
        ELSE
            targetStation := processSequence[sequenceIndex];
            internalState := MOVING;
        END_IF;
END_CASE;

prevSensor1 := sensor1;
prevSensor2 := sensor2;
prevSensor3 := sensor3;
prevSensor4 := sensor4;
prevSensor5 := sensor5;

END_FUNCTION_BLOCK

(* ---- public-hard-02.raw_candidate_01.st ---- *)
FUNCTION_BLOCK FlexibleProcessingControl
VAR_INPUT
    processLength    : USINT;
    sensor1          : BOOL;
    sensor2          : BOOL;
    sensor3          : BOOL;
    sensor4          : BOOL;
    sensor5          : BOOL;
    station1Start    : BOOL;
    station2Complete : BOOL;
    station3Complete : BOOL;
    station4Complete : BOOL;
    processSequence  : ARRAY[1..8] OF USINT;
END_VAR
VAR_OUTPUT
    conveyorLeft  : BOOL;
    conveyorRight : BOOL;
END_VAR
VAR
    state            : INT;
    currentStation   : USINT;
    sequenceIndex    : USINT;
    targetStation    : USINT;
    prevSensor1      : BOOL;
    prevSensor2      : BOOL;
    prevSensor3      : BOOL;
    prevSensor4      : BOOL;
    prevSensor5      : BOOL;
    waitComplete     : BOOL;
END_VAR

(* State constants *)
CONSTANT
    IDLE          : INT := 0;
    LOADING       : INT := 1;
    MOVING        : INT := 2;
    WAIT_PROCESS  : INT := 3;
END_CONSTANT

(* Main logic *)
CASE state OF
    IDLE:
        conveyorLeft  := FALSE;
        conveyorRight := FALSE;
        IF sensor1 AND station1Start THEN
            sequenceIndex  := 1;
            targetStation := processSequence[1];
            currentStation := 1;
            state := LOADING;
        END_IF

    LOADING:
        conveyorLeft  := FALSE;
        conveyorRight := FALSE;
        sequenceIndex := 1;
        targetStation := processSequence[1];
        currentStation := 1;
        state := MOVING;

    MOVING:
        (* Rising edge detection for sensors *)
        IF sensor1 AND NOT prevSensor1 THEN
            currentStation := 1;
        END_IF
        IF sensor2 AND NOT prevSensor2 THEN
            currentStation := 2;
        END_IF
        IF sensor3 AND NOT prevSensor3 THEN
            currentStation := 3;
        END_IF
        IF sensor4 AND NOT prevSensor4 THEN
            currentStation := 4;
        END_IF
        IF sensor5 AND NOT prevSensor5 THEN
            currentStation := 5;
        END_IF

        (* Determine conveyor direction based on target vs current *)
        IF targetStation > currentStation THEN
            conveyorRight := TRUE;
            conveyorLeft  := FALSE;
        ELSIF targetStation < currentStation THEN
            conveyorLeft  := TRUE;
            conveyorRight := FALSE;
        ELSE
            conveyorLeft  := FALSE;
            conveyorRight := FALSE;
        END_IF

        (* Check if product reached target station *)
        IF currentStation = targetStation THEN
            conveyorLeft  := FALSE;
            conveyorRight := FALSE;
            state := WAIT_PROCESS;
            waitComplete := FALSE;
        END_IF

    WAIT_PROCESS:
        IF NOT waitComplete THEN
            waitComplete := TRUE;
        END_IF

        IF waitComplete THEN
            IF targetStation = 2 AND station2Complete THEN
                sequenceIndex := sequenceIndex + 1;
                state := CHECK_SEQUENCE;
            ELSIF targetStation = 3 AND station3Complete THEN
                sequenceIndex := sequenceIndex + 1;
                state := CHECK_SEQUENCE;
            ELSIF targetStation = 4 AND station4Complete THEN
                sequenceIndex := sequenceIndex + 1;
                state := CHECK_SEQUENCE;
            ELSIF targetStation = 5 THEN
                sequenceIndex := sequenceIndex + 1;
                state := CHECK_SEQUENCE;
            END_IF
        END_IF

    CHECK_SEQUENCE:
        IF sequenceIndex > processLength THEN
            state := IDLE;
        ELSE
            targetStation := processSequence[sequenceIndex];
            state := MOVING;
        END_IF
END_CASE

(* Update previous sensor states *)
prevSensor1 := sensor1;
prevSensor2 := sensor2;
prevSensor3 := sensor3;
prevSensor4 := sensor4;
prevSensor5 := sensor5;

END_FUNCTION_BLOCK

(* ---- public-hard-02.raw_candidate_02.st ---- *)
TYPE
    ProcessState : INT (
        IDLE          := 0,
        LOADING       := 1,
        MOVING        := 2,
        WAIT_PROCESS  := 3,
        CHECK_SEQUENCE:= 4
    );
END_TYPE

FUNCTION_BLOCK FlexibleProcessingControl
VAR_INPUT
    processLength    : USINT;
    sensor1          : BOOL;
    sensor2          : BOOL;
    sensor3          : BOOL;
    sensor4          : BOOL;
    sensor5          : BOOL;
    station1Start    : BOOL;
    station2Complete : BOOL;
    station3Complete : BOOL;
    station4Complete : BOOL;
    processSequence  : ARRAY[1..8] OF USINT;
END_VAR
VAR_OUTPUT
    conveyorLeft  : BOOL;
    conveyorRight : BOOL;
END_VAR
VAR
    internalState     : ProcessState;
    currentStation    : USINT;
    sequenceIndex     : USINT;
    targetStation     : USINT;
    prevSensor1       : BOOL;
    prevSensor2       : BOOL;
    prevSensor3       : BOOL;
    prevSensor4       : BOOL;
    prevSensor5       : BOOL;
    waitComplete      : BOOL;
END_VAR

CASE internalState OF
    IDLE:
        conveyorLeft  := FALSE;
        conveyorRight := FALSE;
        IF sensor1 AND station1Start THEN
            sequenceIndex  := 1;
            targetStation := processSequence[1];
            currentStation := 1;
            internalState := LOADING;
        END_IF;

    LOADING:
        conveyorLeft  := FALSE;
        conveyorRight := FALSE;
        sequenceIndex := 1;
        targetStation := processSequence[1];
        currentStation := 1;
        internalState := MOVING;

    MOVING:
        IF sensor1 AND NOT prevSensor1 THEN
            currentStation := 1;
        END_IF;
        IF sensor2 AND NOT prevSensor2 THEN
            currentStation := 2;
        END_IF;
        IF sensor3 AND NOT prevSensor3 THEN
            currentStation := 3;
        END_IF;
        IF sensor4 AND NOT prevSensor4 THEN
            currentStation := 4;
        END_IF;
        IF sensor5 AND NOT prevSensor5 THEN
            currentStation := 5;
        END_IF;

        IF targetStation > currentStation THEN
            conveyorRight := TRUE;
            conveyorLeft  := FALSE;
        ELSIF targetStation < currentStation THEN
            conveyorLeft  := TRUE;
            conveyorRight := FALSE;
        ELSE
            conveyorLeft  := FALSE;
            conveyorRight := FALSE;
        END_IF;

        IF currentStation = targetStation THEN
            conveyorLeft  := FALSE;
            conveyorRight := FALSE;
            internalState := WAIT_PROCESS;
            waitComplete := FALSE;
        END_IF;

    WAIT_PROCESS:
        IF NOT waitComplete THEN
            waitComplete := TRUE;
        END_IF;

        IF waitComplete THEN
            IF targetStation = 2 AND station2Complete THEN
                sequenceIndex := sequenceIndex + 1;
                internalState := CHECK_SEQUENCE;
            ELSIF targetStation = 3 AND station3Complete THEN
                sequenceIndex := sequenceIndex + 1;
                internalState := CHECK_SEQUENCE;
            ELSIF targetStation = 4 AND station4Complete THEN
                sequenceIndex := sequenceIndex + 1;
                internalState := CHECK_SEQUENCE;
            ELSIF targetStation = 5 THEN
                sequenceIndex := sequenceIndex + 1;
                internalState := CHECK_SEQUENCE;
            END_IF;
        END_IF;

    CHECK_SEQUENCE:
        IF sequenceIndex > processLength THEN
            internalState := IDLE;
        ELSE
            targetStation := processSequence[sequenceIndex];
            internalState := MOVING;
        END_IF;
END_CASE;

prevSensor1 := sensor1;
prevSensor2 := sensor2;
prevSensor3 := sensor3;
prevSensor4 := sensor4;
prevSensor5 := sensor5;

END_FUNCTION_BLOCK

(* ---- public-hard-03.candidate_01.st ---- *)
TYPE ST_Recipe :
STRUCT
    recipeID : INT;              (* Recipe identifier; zero denotes an unused database slot. *)
    ingredientType : INT;        (* Ingredient-type identifier. *)
    ingredientRatio : REAL;      (* Ingredient proportion. *)
    productionTemperature : REAL; (* Production temperature. *)
END_STRUCT;
END_TYPE;

FUNCTION_BLOCK RecipeManager
VAR_INPUT
    addRecipe : BOOL;            (* Add Recipe Request Signal *)
    deleteRecipe : BOOL;         (* Delete Recipe Request Signal *)
    modifyRecipe : BOOL;         (* Modify Recipe Request Signal *)
    queryRecipe : BOOL;          (* Query Recipe Request Signal *)
    recipeIn : ST_Recipe;        (* Input Recipe *)
END_VAR

VAR_OUTPUT
    recipeAdded : BOOL;          (* Recipe Added Success Indicator *)
    recipeDeleted : BOOL;        (* Recipe Deleted Success Indicator *)
    recipeModified : BOOL;       (* Recipe Modified Success Indicator *)
    recipeQueryResult : ST_Recipe; (* Recipe Query Result Output *)
    error : BOOL;                (* Error Status Indicator *)
    status : WORD;               (* Status Code *)
END_VAR

VAR_IN_OUT
    recipe : ARRAY[1..10] OF ST_Recipe; (* Recipe Database *)
END_VAR

VAR
    prevAddRecipe : BOOL;
    prevDeleteRecipe : BOOL;
    prevModifyRecipe : BOOL;
    prevQueryRecipe : BOOL;
    i : INT;
    foundIndex : INT;
    emptySlotIndex : INT;
END_VAR

(* Initialize on first cycle *)
IF prevAddRecipe = FALSE AND prevDeleteRecipe = FALSE AND
   prevModifyRecipe = FALSE AND prevQueryRecipe = FALSE THEN
    FOR i := 1 TO 10 DO
        recipe[i].recipeID := 0;
    END_FOR;
END_IF;

(* Clear output flags *)
recipeAdded := FALSE;
recipeDeleted := FALSE;
recipeModified := FALSE;
error := FALSE;
status := 16#0000;

(* Process operations based on rising edge detection *)
IF queryRecipe AND NOT prevQueryRecipe THEN
    foundIndex := 0;
    FOR i := 1 TO 10 DO
        IF recipe[i].recipeID = recipeIn.recipeID THEN
            foundIndex := i;
            EXIT;
        END_IF;
    END_FOR;

    IF foundIndex > 0 THEN
        recipeQueryResult := recipe[foundIndex];
    ELSE
        error := TRUE;
        status := 16#8001;
    END_IF;

ELSIF addRecipe AND NOT prevAddRecipe THEN
    (* Check for duplicate recipeID *)
    foundIndex := 0;
    FOR i := 1 TO 10 DO
        IF recipe[i].recipeID = recipeIn.recipeID THEN
            foundIndex := i;
            EXIT;
        END_IF;
    END_FOR;

    IF foundIndex > 0 THEN
        error := TRUE;
        status := 16#8002;
    ELSE
        (* Find first empty slot *)
        emptySlotIndex := 0;
        FOR i := 1 TO 10 DO
            IF recipe[i].recipeID = 0 THEN
                emptySlotIndex := i;
                EXIT;
            END_IF;
        END_FOR;

        IF emptySlotIndex = 0 THEN
            error := TRUE;
            status := 16#8003;
        ELSE
            recipe[emptySlotIndex] := recipeIn;
            recipeAdded := TRUE;
        END_IF;
    END_IF;

ELSIF deleteRecipe AND NOT prevDeleteRecipe THEN
    foundIndex := 0;
    FOR i := 1 TO 10 DO
        IF recipe[i].recipeID = recipeIn.recipeID THEN
            foundIndex := i;
            EXIT;
        END_IF;
    END_FOR;

    IF foundIndex = 0 THEN
        error := TRUE;
        status := 16#8004;
    ELSE
        recipe[foundIndex].recipeID := 0;
        recipeDeleted := TRUE;
    END_IF;

ELSIF modifyRecipe AND NOT prevModifyRecipe THEN
    foundIndex := 0;
    FOR i := 1 TO 10 DO
        IF recipe[i].recipeID = recipeIn.recipeID THEN
            foundIndex := i;
            EXIT;
        END_IF;
    END_FOR;

    IF foundIndex = 0 THEN
        error := TRUE;
        status := 16#8005;
    ELSE
        recipe[foundIndex] := recipeIn;
        recipeModified := TRUE;
    END_IF;
END_IF;

(* Update edge detection state *)
prevAddRecipe := addRecipe;
prevDeleteRecipe := deleteRecipe;
prevModifyRecipe := modifyRecipe;
prevQueryRecipe := queryRecipe;

END_FUNCTION_BLOCK

(* ---- public-hard-03.candidate_02.st ---- *)
TYPE ST_Recipe :
STRUCT
    recipeID : INT
    ingredientType : INT
    ingredientRatio : REAL
    productionTemperature : REAL
END_STRUCT;
END_TYPE;

FUNCTION_BLOCK RecipeManager
VAR_INPUT
    addRecipe : BOOL;
    deleteRecipe : BOOL;
    modifyRecipe : BOOL;
    queryRecipe : BOOL;
    recipeIn : ST_Recipe;
END_VAR

VAR_OUTPUT
    recipeAdded : BOOL;
    recipeDeleted : BOOL;
    recipeModified : BOOL;
    recipeQueryResult : ST_Recipe;
    error : BOOL;
    status : WORD;
END_VAR

VAR_IN_OUT
    recipe : ARRAY[1..10] OF ST_Recipe;
END_VAR

VAR
    prevAddRecipe : BOOL;
    prevDeleteRecipe : BOOL;
    prevModifyRecipe : BOOL;
    prevQueryRecipe : BOOL;
    i : INT;
    foundIndex : INT;
    emptySlotIndex : INT;
END_VAR

IF prevAddRecipe = FALSE AND prevDeleteRecipe = FALSE AND
   prevModifyRecipe = FALSE AND prevQueryRecipe = FALSE THEN
    FOR i := 1 TO 10 DO
        recipe[i].recipeID := 0;
    END_FOR;
END_IF;

recipeAdded := FALSE;
recipeDeleted := FALSE;
recipeModified := FALSE;
error := FALSE;
status := 16#0000;

IF queryRecipe AND NOT prevQueryRecipe THEN
    foundIndex := 0;
    FOR i := 1 TO 10 DO
        IF recipe[i].recipeID = recipeIn.recipeID THEN
            foundIndex := i;
            EXIT;
        END_IF;
    END_FOR;

    IF foundIndex > 0 THEN
        recipeQueryResult := recipe[foundIndex];
    ELSE
        error := TRUE;
        status := 16#8001;
    END_IF;

ELSIF addRecipe AND NOT prevAddRecipe THEN
    foundIndex := 0;
    FOR i := 1 TO 10 DO
        IF recipe[i].recipeID = recipeIn.recipeID THEN
            foundIndex := i;
            EXIT;
        END_IF;
    END_FOR;

    IF foundIndex > 0 THEN
        error := TRUE;
        status := 16#8002;
    ELSE
        emptySlotIndex := 0;
        FOR i := 1 TO 10 DO
            IF recipe[i].recipeID = 0 THEN
                emptySlotIndex := i;
                EXIT;
            END_IF;
        END_FOR;

        IF emptySlotIndex = 0 THEN
            error := TRUE;
            status := 16#8003;
        ELSE
            recipe[emptySlotIndex] := recipeIn;
            recipeAdded := TRUE;
        END_IF;
    END_IF;

ELSIF deleteRecipe AND NOT prevDeleteRecipe THEN
    foundIndex := 0;
    FOR i := 1 TO 10 DO
        IF recipe[i].recipeID = recipeIn.recipeID THEN
            foundIndex := i;
            EXIT;
        END_IF;
    END_FOR;

    IF foundIndex = 0 THEN
        error := TRUE;
        status := 16#8004;
    ELSE
        recipe[foundIndex].recipeID := 0;
        recipeDeleted := TRUE;
    END_IF;

ELSIF modifyRecipe AND NOT prevModifyRecipe THEN
    foundIndex := 0;
    FOR i := 1 TO 10 DO
        IF recipe[i].recipeID = recipeIn.recipeID THEN
            foundIndex := i;
            EXIT;
        END_IF;
    END_FOR;

    IF foundIndex = 0 THEN
        error := TRUE;
        status := 16#8005;
    ELSE
        recipe[foundIndex] := recipeIn;
        recipeModified := TRUE;
    END_IF;
END_IF;

prevAddRecipe := addRecipe;
prevDeleteRecipe := deleteRecipe;
prevModifyRecipe := modifyRecipe;
prevQueryRecipe := queryRecipe;

END_FUNCTION_BLOCK

(* ---- public-hard-03.raw_candidate_01.st ---- *)
TYPE ST_Recipe :
STRUCT
    recipeID : INT;              (* Recipe identifier; zero denotes an unused database slot. *)
    ingredientType : INT;        (* Ingredient-type identifier. *)
    ingredientRatio : REAL;      (* Ingredient proportion. *)
    productionTemperature : REAL; (* Production temperature. *)
END_STRUCT
END_TYPE

FUNCTION_BLOCK RecipeManager
VAR_INPUT
    addRecipe : BOOL;            (* Add Recipe Request Signal *)
    deleteRecipe : BOOL;         (* Delete Recipe Request Signal *)
    modifyRecipe : BOOL;         (* Modify Recipe Request Signal *)
    queryRecipe : BOOL;          (* Query Recipe Request Signal *)
    recipeIn : ST_Recipe;        (* Input Recipe *)
END_VAR

VAR_OUTPUT
    recipeAdded : BOOL;          (* Recipe Added Success Indicator *)
    recipeDeleted : BOOL;        (* Recipe Deleted Success Indicator *)
    recipeModified : BOOL;       (* Recipe Modified Success Indicator *)
    recipeQueryResult : ST_Recipe; (* Recipe Query Result Output *)
    error : BOOL;                (* Error Status Indicator *)
    status : WORD;               (* Status Code *)
END_VAR

VAR_IN_OUT
    recipe : ARRAY[1..10] OF ST_Recipe; (* Recipe Database *)
END_VAR

VAR
    prevAddRecipe : BOOL;
    prevDeleteRecipe : BOOL;
    prevModifyRecipe : BOOL;
    prevQueryRecipe : BOOL;
    i : INT;
    foundIndex : INT;
    emptySlotIndex : INT;
END_VAR

(* Initialize on first cycle *)
IF prevAddRecipe = FALSE AND prevDeleteRecipe = FALSE AND
   prevModifyRecipe = FALSE AND prevQueryRecipe = FALSE THEN
    FOR i := 1 TO 10 DO
        recipe[i].recipeID := 0;
    END_FOR;
END_IF;

(* Clear output flags *)
recipeAdded := FALSE;
recipeDeleted := FALSE;
recipeModified := FALSE;
error := FALSE;
status := 16#0000;

(* Process operations based on rising edge detection *)
IF queryRecipe AND NOT prevQueryRecipe THEN
    foundIndex := 0;
    FOR i := 1 TO 10 DO
        IF recipe[i].recipeID = recipeIn.recipeID THEN
            foundIndex := i;
            EXIT;
        END_IF;
    END_FOR;

    IF foundIndex > 0 THEN
        recipeQueryResult := recipe[foundIndex];
    ELSE
        error := TRUE;
        status := 16#8001;
    END_IF;

ELSIF addRecipe AND NOT prevAddRecipe THEN
    (* Check for duplicate recipeID *)
    foundIndex := 0;
    FOR i := 1 TO 10 DO
        IF recipe[i].recipeID = recipeIn.recipeID THEN
            foundIndex := i;
            EXIT;
        END_IF;
    END_FOR;

    IF foundIndex > 0 THEN
        error := TRUE;
        status := 16#8002;
    ELSE
        (* Find first empty slot *)
        emptySlotIndex := 0;
        FOR i := 1 TO 10 DO
            IF recipe[i].recipeID = 0 THEN
                emptySlotIndex := i;
                EXIT;
            END_IF;
        END_FOR;

        IF emptySlotIndex = 0 THEN
            error := TRUE;
            status := 16#8003;
        ELSE
            recipe[emptySlotIndex] := recipeIn;
            recipeAdded := TRUE;
        END_IF;
    END_IF;

ELSIF deleteRecipe AND NOT prevDeleteRecipe THEN
    foundIndex := 0;
    FOR i := 1 TO 10 DO
        IF recipe[i].recipeID = recipeIn.recipeID THEN
            foundIndex := i;
            EXIT;
        END_IF;
    END_FOR;

    IF foundIndex = 0 THEN
        error := TRUE;
        status := 16#8004;
    ELSE
        recipe[foundIndex].recipeID := 0;
        recipeDeleted := TRUE;
    END_IF;

ELSIF modifyRecipe AND NOT prevModifyRecipe THEN
    foundIndex := 0;
    FOR i := 1 TO 10 DO
        IF recipe[i].recipeID = recipeIn.recipeID THEN
            foundIndex := i;
            EXIT;
        END_IF;
    END_FOR;

    IF foundIndex = 0 THEN
        error := TRUE;
        status := 16#8005;
    ELSE
        recipe[foundIndex] := recipeIn;
        recipeModified := TRUE;
    END_IF;
END_IF;

(* Update edge detection state *)
prevAddRecipe := addRecipe;
prevDeleteRecipe := deleteRecipe;
prevModifyRecipe := modifyRecipe;
prevQueryRecipe := queryRecipe;

END_FUNCTION_BLOCK

(* ---- public-hard-03.raw_candidate_02.st ---- *)
TYPE ST_Recipe :
STRUCT
    recipeID : INT
    ingredientType : INT
    ingredientRatio : REAL
    productionTemperature : REAL
END_STRUCT
END_TYPE

FUNCTION_BLOCK RecipeManager
VAR_INPUT
    addRecipe : BOOL;
    deleteRecipe : BOOL;
    modifyRecipe : BOOL;
    queryRecipe : BOOL;
    recipeIn : ST_Recipe;
END_VAR

VAR_OUTPUT
    recipeAdded : BOOL;
    recipeDeleted : BOOL;
    recipeModified : BOOL;
    recipeQueryResult : ST_Recipe;
    error : BOOL;
    status : WORD;
END_VAR

VAR_IN_OUT
    recipe : ARRAY[1..10] OF ST_Recipe;
END_VAR

VAR
    prevAddRecipe : BOOL;
    prevDeleteRecipe : BOOL;
    prevModifyRecipe : BOOL;
    prevQueryRecipe : BOOL;
    i : INT;
    foundIndex : INT;
    emptySlotIndex : INT;
END_VAR

IF prevAddRecipe = FALSE AND prevDeleteRecipe = FALSE AND
   prevModifyRecipe = FALSE AND prevQueryRecipe = FALSE THEN
    FOR i := 1 TO 10 DO
        recipe[i].recipeID := 0;
    END_FOR;
END_IF;

recipeAdded := FALSE;
recipeDeleted := FALSE;
recipeModified := FALSE;
error := FALSE;
status := 16#0000;

IF queryRecipe AND NOT prevQueryRecipe THEN
    foundIndex := 0;
    FOR i := 1 TO 10 DO
        IF recipe[i].recipeID = recipeIn.recipeID THEN
            foundIndex := i;
            EXIT;
        END_IF;
    END_FOR;

    IF foundIndex > 0 THEN
        recipeQueryResult := recipe[foundIndex];
    ELSE
        error := TRUE;
        status := 16#8001;
    END_IF;

ELSIF addRecipe AND NOT prevAddRecipe THEN
    foundIndex := 0;
    FOR i := 1 TO 10 DO
        IF recipe[i].recipeID = recipeIn.recipeID THEN
            foundIndex := i;
            EXIT;
        END_IF;
    END_FOR;

    IF foundIndex > 0 THEN
        error := TRUE;
        status := 16#8002;
    ELSE
        emptySlotIndex := 0;
        FOR i := 1 TO 10 DO
            IF recipe[i].recipeID = 0 THEN
                emptySlotIndex := i;
                EXIT;
            END_IF;
        END_FOR;

        IF emptySlotIndex = 0 THEN
            error := TRUE;
            status := 16#8003;
        ELSE
            recipe[emptySlotIndex] := recipeIn;
            recipeAdded := TRUE;
        END_IF;
    END_IF;

ELSIF deleteRecipe AND NOT prevDeleteRecipe THEN
    foundIndex := 0;
    FOR i := 1 TO 10 DO
        IF recipe[i].recipeID = recipeIn.recipeID THEN
            foundIndex := i;
            EXIT;
        END_IF;
    END_FOR;

    IF foundIndex = 0 THEN
        error := TRUE;
        status := 16#8004;
    ELSE
        recipe[foundIndex].recipeID := 0;
        recipeDeleted := TRUE;
    END_IF;

ELSIF modifyRecipe AND NOT prevModifyRecipe THEN
    foundIndex := 0;
    FOR i := 1 TO 10 DO
        IF recipe[i].recipeID = recipeIn.recipeID THEN
            foundIndex := i;
            EXIT;
        END_IF;
    END_FOR;

    IF foundIndex = 0 THEN
        error := TRUE;
        status := 16#8005;
    ELSE
        recipe[foundIndex] := recipeIn;
        recipeModified := TRUE;
    END_IF;
END_IF;

prevAddRecipe := addRecipe;
prevDeleteRecipe := deleteRecipe;
prevModifyRecipe := modifyRecipe;
prevQueryRecipe := queryRecipe;

END_FUNCTION_BLOCK

(* ---- public-hard-04.candidate_01.st ---- *)
FUNCTION_BLOCK FB_FIFOQueue
VAR_INPUT
    enqueue : BOOL;
    dequeue : BOOL;
    reset   : BOOL;
END_VAR
VAR_OUTPUT
    elementCount : DINT;
    status       : WORD;
END_VAR
VAR_IN_OUT
    item   : VARIANT;
    buffer : VARIANT;
END_VAR
VAR
    head        : DINT := 0;
    tail        : DINT := 0;
    capacity    : DINT := 0;
    prevEnqueue : BOOL := FALSE;
    prevDequeue : BOOL := FALSE;
    prevReset   : BOOL := FALSE;
END_VAR

status := 16#0000;

IF reset AND NOT prevReset THEN
    head := 0;
    tail := 0;
    elementCount := 0;
ELSIF enqueue AND NOT prevEnqueue THEN
    IF capacity > 0 AND elementCount < capacity THEN
        buffer[tail] := item;
        tail := (tail + 1) MOD capacity;
        elementCount := elementCount + 1;
    ELSIF elementCount >= capacity THEN
        status := 16#8002;
    END_IF;
ELSIF dequeue AND NOT prevDequeue THEN
    IF elementCount > 0 THEN
        item := buffer[head];
        head := (head + 1) MOD capacity;
        elementCount := elementCount - 1;
    ELSE
        status := 16#8001;
    END_IF;
END_IF;

IF capacity = 0 AND __ISARRAY(buffer) THEN
    capacity := __UPPERBOUND(buffer, 1) - __LOWERBOUND(buffer, 1) + 1;
END_IF;

prevEnqueue := enqueue;
prevDequeue := dequeue;
prevReset := reset;
END_FUNCTION_BLOCK

(* ---- public-hard-04.candidate_02.st ---- *)
FUNCTION_BLOCK FB_FIFOQueue
VAR_INPUT
    enqueue : BOOL;
    dequeue : BOOL;
    reset   : BOOL;
END_VAR
VAR_OUTPUT
    elementCount : DINT;
    status       : WORD;
END_VAR
VAR_IN_OUT
    item   : VARIANT;
    buffer : VARIANT;
END_VAR
VAR
    head       : DINT := 0;
    tail       : DINT := 0;
    capacity   : DINT := 0;
    prevEnqueue : BOOL := FALSE;
    prevDequeue : BOOL := FALSE;
    prevReset   : BOOL := FALSE;
    firstCall   : BOOL := TRUE;
END_VAR

status := 16#0000;

IF firstCall THEN
    firstCall := FALSE;
    prevEnqueue := enqueue;
    prevDequeue := dequeue;
    prevReset := reset;
    RETURN;
END_IF;

IF __ISARRAY(buffer) THEN
    capacity := __UBOUND(buffer, 1) - __LBBOUND(buffer, 1) + 1;
END_IF;

IF reset AND NOT prevReset THEN
    head := 0;
    tail := 0;
    elementCount := 0;
ELSIF enqueue AND NOT prevEnqueue THEN
    IF elementCount < capacity THEN
        buffer[tail] := item;
        tail := (tail + 1) MOD capacity;
        elementCount := elementCount + 1;
    ELSE
        status := 16#8002;
    END_IF;
ELSIF dequeue AND NOT prevDequeue THEN
    IF elementCount > 0 THEN
        item := buffer[head];
        head := (head + 1) MOD capacity;
        elementCount := elementCount - 1;
    ELSE
        status := 16#8001;
    END_IF;
END_IF;

prevEnqueue := enqueue;
prevDequeue := dequeue;
prevReset := reset;
END_FUNCTION_BLOCK

(* ---- public-hard-04.raw_candidate_01.st ---- *)
FUNCTION_BLOCK FB_FIFOQueue
VAR_INPUT
    enqueue : BOOL;
    dequeue : BOOL;
    reset   : BOOL;
END_VAR
VAR_OUTPUT
    elementCount : DINT;
    status       : WORD;
END_VAR
VAR_IN_OUT
    item   : VARIANT;
    buffer : VARIANT;
END_VAR
VAR
    head        : DINT := 0;
    tail        : DINT := 0;
    capacity    : DINT := 0;
    prevEnqueue : BOOL := FALSE;
    prevDequeue : BOOL := FALSE;
    prevReset   : BOOL := FALSE;
END_VAR

status := 16#0000;

IF reset AND NOT prevReset THEN
    head := 0;
    tail := 0;
    elementCount := 0;
ELSIF enqueue AND NOT prevEnqueue THEN
    IF capacity > 0 AND elementCount < capacity THEN
        buffer[tail] := item;
        tail := (tail + 1) MOD capacity;
        elementCount := elementCount + 1;
    ELSIF elementCount >= capacity THEN
        status := 16#8002;
    END_IF;
ELSIF dequeue AND NOT prevDequeue THEN
    IF elementCount > 0 THEN
        item := buffer[head];
        head := (head + 1) MOD capacity;
        elementCount := elementCount - 1;
    ELSE
        status := 16#8001;
    END_IF;
END_IF;

IF capacity = 0 AND __ISARRAY(buffer) THEN
    capacity := __UPPERBOUND(buffer, 1) - __LOWERBOUND(buffer, 1) + 1;
END_IF;

prevEnqueue := enqueue;
prevDequeue := dequeue;
prevReset := reset;
END_FUNCTION_BLOCK

(* ---- public-hard-04.raw_candidate_02.st ---- *)
FUNCTION_BLOCK FB_FIFOQueue
VAR_INPUT
    enqueue : BOOL;
    dequeue : BOOL;
    reset   : BOOL;
END_VAR
VAR_OUTPUT
    elementCount : DINT;
    status       : WORD;
END_VAR
VAR_IN_OUT
    item   : VARIANT;
    buffer : VARIANT;
END_VAR
VAR
    head       : DINT := 0;
    tail       : DINT := 0;
    capacity   : DINT := 0;
    prevEnqueue : BOOL := FALSE;
    prevDequeue : BOOL := FALSE;
    prevReset   : BOOL := FALSE;
    firstCall   : BOOL := TRUE;
END_VAR

status := 16#0000;

IF firstCall THEN
    firstCall := FALSE;
    prevEnqueue := enqueue;
    prevDequeue := dequeue;
    prevReset := reset;
    RETURN;
END_IF

IF __ISARRAY(buffer) THEN
    capacity := __UBOUND(buffer, 1) - __LBBOUND(buffer, 1) + 1;
END_IF;

IF reset AND NOT prevReset THEN
    head := 0;
    tail := 0;
    elementCount := 0;
ELSIF enqueue AND NOT prevEnqueue THEN
    IF elementCount < capacity THEN
        buffer[tail] := item;
        tail := (tail + 1) MOD capacity;
        elementCount := elementCount + 1;
    ELSE
        status := 16#8002;
    END_IF;
ELSIF dequeue AND NOT prevDequeue THEN
    IF elementCount > 0 THEN
        item := buffer[head];
        head := (head + 1) MOD capacity;
        elementCount := elementCount - 1;
    ELSE
        status := 16#8001;
    END_IF;
END_IF;

prevEnqueue := enqueue;
prevDequeue := dequeue;
prevReset := reset;
END_FUNCTION_BLOCK

(* ---- public-hard-05.candidate_01.st ---- *)
FUNCTION_BLOCK MechanicalArmControl
VAR_INPUT
    ManualMode      : BOOL;
    SingleStepMode  : BOOL;
    SingleCycleMode : BOOL;
    ContinuousMode  : BOOL;
    EmergencyStop   : BOOL;
    Start           : BOOL;
    DownButton      : BOOL;
    UpButton        : BOOL;
    LeftButton      : BOOL;
    RightButton     : BOOL;
    GripButton      : BOOL;
    ReleaseButton   : BOOL;
    DownLimitSwitch     : BOOL;
    UpLimitSwitch       : BOOL;
    LeftLimitSwitch     : BOOL;
    RightLimitSwitch    : BOOL;
    GripLimitSwitch     : BOOL;
    ReleaseLimitSwitch  : BOOL;
END_VAR

VAR_OUTPUT
    MoveDown        : BOOL;
    MoveUp          : BOOL;
    MoveLeft        : BOOL;
    MoveRight       : BOOL;
    ActivateGrip    : BOOL;
    ActivateRelease : BOOL;
END_VAR

VAR
    stepNumber       : INT := 0;
    startRisingEdge  : BOOL;
    lastStart        : BOOL := FALSE;
    actionInProgress : BOOL := FALSE;
END_VAR

// Edge detection for Start button
startRisingEdge := Start AND NOT lastStart;
lastStart := Start;

// Emergency stop: highest priority, resets all outputs and state
IF NOT EmergencyStop THEN
    MoveDown        := FALSE;
    MoveUp          := FALSE;
    MoveLeft        := FALSE;
    MoveRight       := FALSE;
    ActivateGrip    := FALSE;
    ActivateRelease := FALSE;
    stepNumber      := 0;
    actionInProgress := FALSE;
ELSE
    // Manual mode control
    IF ManualMode THEN
        MoveDown        := DownButton AND NOT DownLimitSwitch;
        MoveUp          := UpButton AND NOT UpLimitSwitch;
        MoveLeft        := LeftButton AND NOT LeftLimitSwitch;
        MoveRight       := RightButton AND NOT RightLimitSwitch;
        ActivateGrip    := GripButton AND NOT GripLimitSwitch;
        ActivateRelease := ReleaseButton AND NOT ReleaseLimitSwitch;
        stepNumber      := 0;
        actionInProgress := FALSE;

    // Single step mode: Start button advances through steps
    ELSIF SingleStepMode THEN
        IF startRisingEdge AND NOT actionInProgress THEN
            stepNumber := stepNumber + 1;
        END_IF;

        CASE stepNumber OF
            1:
                MoveDown := TRUE;
                actionInProgress := TRUE;
                IF DownLimitSwitch THEN
                    MoveDown := FALSE;
                    actionInProgress := FALSE;
                END_IF;
            2:
                ActivateGrip := TRUE;
                actionInProgress := TRUE;
                IF GripLimitSwitch THEN
                    ActivateGrip := FALSE;
                    actionInProgress := FALSE;
                END_IF;
            3:
                MoveUp := TRUE;
                actionInProgress := TRUE;
                IF UpLimitSwitch THEN
                    MoveUp := FALSE;
                    actionInProgress := FALSE;
                END_IF;
            4:
                MoveRight := TRUE;
                actionInProgress := TRUE;
                IF RightLimitSwitch THEN
                    MoveRight := FALSE;
                    actionInProgress := FALSE;
                END_IF;
            5:
                MoveDown := TRUE;
                actionInProgress := TRUE;
                IF DownLimitSwitch THEN
                    MoveDown := FALSE;
                    actionInProgress := FALSE;
                END_IF;
            6:
                ActivateRelease := TRUE;
                actionInProgress := TRUE;
                IF ReleaseLimitSwitch THEN
                    ActivateRelease := FALSE;
                    actionInProgress := FALSE;
                END_IF;
            7:
                MoveUp := TRUE;
                actionInProgress := TRUE;
                IF UpLimitSwitch THEN
                    MoveUp := FALSE;
                    actionInProgress := FALSE;
                END_IF;
            8:
                MoveLeft := TRUE;
                actionInProgress := TRUE;
                IF LeftLimitSwitch THEN
                    MoveLeft := FALSE;
                    actionInProgress := FALSE;
                END_IF;
        END_CASE;

        IF stepNumber > 8 THEN
            stepNumber := 0;
        END_IF;

    // Single cycle mode: executes full cycle once then stops
    ELSIF SingleCycleMode THEN
        IF startRisingEdge THEN
            stepNumber := 1;
            actionInProgress := FALSE;
        END_IF;

        CASE stepNumber OF
            1:
                MoveDown := TRUE;
                actionInProgress := TRUE;
                IF DownLimitSwitch THEN
                    MoveDown := FALSE;
                    actionInProgress := FALSE;
                    stepNumber := 2;
                END_IF;
            2:
                ActivateGrip := TRUE;
                actionInProgress := TRUE;
                IF GripLimitSwitch THEN
                    ActivateGrip := FALSE;
                    actionInProgress := FALSE;
                    stepNumber := 3;
                END_IF;
            3:
                MoveUp := TRUE;
                actionInProgress := TRUE;
                IF UpLimitSwitch THEN
                    MoveUp := FALSE;
                    actionInProgress := FALSE;
                    stepNumber := 4;
                END_IF;
            4:
                MoveRight := TRUE;
                actionInProgress := TRUE;
                IF RightLimitSwitch THEN
                    MoveRight := FALSE;
                    actionInProgress := FALSE;
                    stepNumber := 5;
                END_IF;
            5:
                MoveDown := TRUE;
                actionInProgress := TRUE;
                IF DownLimitSwitch THEN
                    MoveDown := FALSE;
                    actionInProgress := FALSE;
                    stepNumber := 6;
                END_IF;
            6:
                ActivateRelease := TRUE;
                actionInProgress := TRUE;
                IF ReleaseLimitSwitch THEN
                    ActivateRelease := FALSE;
                    actionInProgress := FALSE;
                    stepNumber := 7;
                END_IF;
            7:
                MoveUp := TRUE;
                actionInProgress := TRUE;
                IF UpLimitSwitch THEN
                    MoveUp := FALSE;
                    actionInProgress := FALSE;
                    stepNumber := 8;
                END_IF;
            8:
                MoveLeft := TRUE;
                actionInProgress := TRUE;
                IF LeftLimitSwitch THEN
                    MoveLeft := FALSE;
                    actionInProgress := FALSE;
                    stepNumber := 0;
                END_IF;
        END_CASE;

    // Continuous mode: executes full cycle repeatedly
    ELSIF ContinuousMode THEN
        IF startRisingEdge THEN
            stepNumber := 1;
            actionInProgress := FALSE;
        END_IF;

        CASE stepNumber OF
            1:
                MoveDown := TRUE;
                actionInProgress := TRUE;
                IF DownLimitSwitch THEN
                    MoveDown := FALSE;
                    actionInProgress := FALSE;
                    stepNumber := 2;
                END_IF;
            2:
                ActivateGrip := TRUE;
                actionInProgress := TRUE;
                IF GripLimitSwitch THEN
                    ActivateGrip := FALSE;
                    actionInProgress := FALSE;
                    stepNumber := 3;
                END_IF;
            3:
                MoveUp := TRUE;
                actionInProgress := TRUE;
                IF UpLimitSwitch THEN
                    MoveUp := FALSE;
                    actionInProgress := FALSE;
                    stepNumber := 4;
                END_IF;
            4:
                MoveRight := TRUE;
                actionInProgress := TRUE;
                IF RightLimitSwitch THEN
                    MoveRight := FALSE;
                    actionInProgress := FALSE;
                    stepNumber := 5;
                END_IF;
            5:
                MoveDown := TRUE;
                actionInProgress := TRUE;
                IF DownLimitSwitch THEN
                    MoveDown := FALSE;
                    actionInProgress := FALSE;
                    stepNumber := 6;
                END_IF;
            6:
                ActivateRelease := TRUE;
                actionInProgress := TRUE;
                IF ReleaseLimitSwitch THEN
                    ActivateRelease := FALSE;
                    actionInProgress := FALSE;
                    stepNumber := 7;
                END_IF;
            7:
                MoveUp := TRUE;
                actionInProgress := TRUE;
                IF UpLimitSwitch THEN
                    MoveUp := FALSE;
                    actionInProgress := FALSE;
                    stepNumber := 8;
                END_IF;
            8:
                MoveLeft := TRUE;
                actionInProgress := TRUE;
                IF LeftLimitSwitch THEN
                    MoveLeft := FALSE;
                    actionInProgress := FALSE;
                    stepNumber := 1;
                END_IF;
        END_CASE;
    END_IF;
END_IF;
END_FUNCTION_BLOCK

(* ---- public-hard-05.candidate_02.st ---- *)
FUNCTION_BLOCK MechanicalArmControl
VAR_INPUT
    ManualMode      : BOOL;
    SingleStepMode  : BOOL;
    SingleCycleMode : BOOL;
    ContinuousMode  : BOOL;
    EmergencyStop   : BOOL;
    Start           : BOOL;
    DownButton      : BOOL;
    UpButton        : BOOL;
    LeftButton      : BOOL;
    RightButton     : BOOL;
    GripButton      : BOOL;
    ReleaseButton   : BOOL;
    DownLimitSwitch     : BOOL;
    UpLimitSwitch       : BOOL;
    LeftLimitSwitch     : BOOL;
    RightLimitSwitch    : BOOL;
    GripLimitSwitch     : BOOL;
    ReleaseLimitSwitch  : BOOL;
END_VAR

VAR_OUTPUT
    MoveDown        : BOOL;
    MoveUp          : BOOL;
    MoveLeft        : BOOL;
    MoveRight       : BOOL;
    ActivateGrip    : BOOL;
    ActivateRelease : BOOL;
END_VAR

VAR
    stepNumber       : INT := 0;
    startRisingEdge  : BOOL;
    lastStart        : BOOL := FALSE;
    actionInProgress : BOOL := FALSE;
END_VAR

startRisingEdge := Start AND NOT lastStart;
lastStart := Start;

IF NOT EmergencyStop THEN
    MoveDown        := FALSE;
    MoveUp          := FALSE;
    MoveLeft        := FALSE;
    MoveRight       := FALSE;
    ActivateGrip    := FALSE;
    ActivateRelease := FALSE;
    stepNumber      := 0;
    actionInProgress := FALSE;
ELSE
    IF ManualMode THEN
        IF DownButton AND UpButton THEN
            MoveDown := FALSE;
            MoveUp := FALSE;
        ELSE
            MoveDown := DownButton AND NOT DownLimitSwitch;
            MoveUp := UpButton AND NOT UpLimitSwitch;
        END_IF;
        IF LeftButton AND RightButton THEN
            MoveLeft := FALSE;
            MoveRight := FALSE;
        ELSE
            MoveLeft := LeftButton AND NOT LeftLimitSwitch;
            MoveRight := RightButton AND NOT RightLimitSwitch;
        END_IF;
        ActivateGrip := GripButton AND NOT GripLimitSwitch;
        ActivateRelease := ReleaseButton AND NOT ReleaseLimitSwitch;
        stepNumber := 0;
        actionInProgress := FALSE;

    ELSIF SingleStepMode THEN
        IF startRisingEdge AND NOT actionInProgress THEN
            stepNumber := stepNumber + 1;
        END_IF;

        IF stepNumber = 0 THEN
            actionInProgress := FALSE;
        END_IF;

        CASE stepNumber OF
            1:
                MoveDown := TRUE;
                actionInProgress := TRUE;
                IF DownLimitSwitch THEN
                    MoveDown := FALSE;
                    actionInProgress := FALSE;
                END_IF;
            2:
                ActivateGrip := TRUE;
                actionInProgress := TRUE;
                IF GripLimitSwitch THEN
                    ActivateGrip := FALSE;
                    actionInProgress := FALSE;
                END_IF;
            3:
                MoveUp := TRUE;
                actionInProgress := TRUE;
                IF UpLimitSwitch THEN
                    MoveUp := FALSE;
                    actionInProgress := FALSE;
                END_IF;
            4:
                MoveRight := TRUE;
                actionInProgress := TRUE;
                IF RightLimitSwitch THEN
                    MoveRight := FALSE;
                    actionInProgress := FALSE;
                END_IF;
            5:
                MoveDown := TRUE;
                actionInProgress := TRUE;
                IF DownLimitSwitch THEN
                    MoveDown := FALSE;
                    actionInProgress := FALSE;
                END_IF;
            6:
                ActivateRelease := TRUE;
                actionInProgress := TRUE;
                IF ReleaseLimitSwitch THEN
                    ActivateRelease := FALSE;
                    actionInProgress := FALSE;
                END_IF;
            7:
                MoveUp := TRUE;
                actionInProgress := TRUE;
                IF UpLimitSwitch THEN
                    MoveUp := FALSE;
                    actionInProgress := FALSE;
                END_IF;
            8:
                MoveLeft := TRUE;
                actionInProgress := TRUE;
                IF LeftLimitSwitch THEN
                    MoveLeft := FALSE;
                    actionInProgress := FALSE;
                END_IF;
        END_CASE;

        IF stepNumber > 8 THEN
            stepNumber := 0;
        END_IF;

    ELSIF SingleCycleMode THEN
        IF startRisingEdge THEN
            stepNumber := 1;
            actionInProgress := FALSE;
        END_IF;

        IF stepNumber = 0 THEN
            actionInProgress := FALSE;
        END_IF;

        CASE stepNumber OF
            1:
                MoveDown := TRUE;
                actionInProgress := TRUE;
                IF DownLimitSwitch THEN
                    MoveDown := FALSE;
                    actionInProgress := FALSE;
                    stepNumber := 2;
                END_IF;
            2:
                ActivateGrip := TRUE;
                actionInProgress := TRUE;
                IF GripLimitSwitch THEN
                    ActivateGrip := FALSE;
                    actionInProgress := FALSE;
                    stepNumber := 3;
                END_IF;
            3:
                MoveUp := TRUE;
                actionInProgress := TRUE;
                IF UpLimitSwitch THEN
                    MoveUp := FALSE;
                    actionInProgress := FALSE;
                    stepNumber := 4;
                END_IF;
            4:
                MoveRight := TRUE;
                actionInProgress := TRUE;
                IF RightLimitSwitch THEN
                    MoveRight := FALSE;
                    actionInProgress := FALSE;
                    stepNumber := 5;
                END_IF;
            5:
                MoveDown := TRUE;
                actionInProgress := TRUE;
                IF DownLimitSwitch THEN
                    MoveDown := FALSE;
                    actionInProgress := FALSE;
                    stepNumber := 6;
                END_IF;
            6:
                ActivateRelease := TRUE;
                actionInProgress := TRUE;
                IF ReleaseLimitSwitch THEN
                    ActivateRelease := FALSE;
                    actionInProgress := FALSE;
                    stepNumber := 7;
                END_IF;
            7:
                MoveUp := TRUE;
                actionInProgress := TRUE;
                IF UpLimitSwitch THEN
                    MoveUp := FALSE;
                    actionInProgress := FALSE;
                    stepNumber := 8;
                END_IF;
            8:
                MoveLeft := TRUE;
                actionInProgress := TRUE;
                IF LeftLimitSwitch THEN
                    MoveLeft := FALSE;
                    actionInProgress := FALSE;
                    stepNumber := 0;
                END_IF;
        END_CASE;

    ELSIF ContinuousMode THEN
        IF startRisingEdge THEN
            stepNumber := 1;
            actionInProgress := FALSE;
        END_IF;

        IF stepNumber = 0 THEN
            actionInProgress := FALSE;
        END_IF;

        CASE stepNumber OF
            1:
                MoveDown := TRUE;
                actionInProgress := TRUE;
                IF DownLimitSwitch THEN
                    MoveDown := FALSE;
                    actionInProgress := FALSE;
                    stepNumber := 2;
                END_IF;
            2:
                ActivateGrip := TRUE;
                actionInProgress := TRUE;
                IF GripLimitSwitch THEN
                    ActivateGrip := FALSE;
                    actionInProgress := FALSE;
                    stepNumber := 3;
                END_IF;
            3:
                MoveUp := TRUE;
                actionInProgress := TRUE;
                IF UpLimitSwitch THEN
                    MoveUp := FALSE;
                    actionInProgress := FALSE;
                    stepNumber := 4;
                END_IF;
            4:
                MoveRight := TRUE;
                actionInProgress := TRUE;
                IF RightLimitSwitch THEN
                    MoveRight := FALSE;
                    actionInProgress := FALSE;
                    stepNumber := 5;
                END_IF;
            5:
                MoveDown := TRUE;
                actionInProgress := TRUE;
                IF DownLimitSwitch THEN
                    MoveDown := FALSE;
                    actionInProgress := FALSE;
                    stepNumber := 6;
                END_IF;
            6:
                ActivateRelease := TRUE;
                actionInProgress := TRUE;
                IF ReleaseLimitSwitch THEN
                    ActivateRelease := FALSE;
                    actionInProgress := FALSE;
                    stepNumber := 7;
                END_IF;
            7:
                MoveUp := TRUE;
                actionInProgress := TRUE;
                IF UpLimitSwitch THEN
                    MoveUp := FALSE;
                    actionInProgress := FALSE;
                    stepNumber := 8;
                END_IF;
            8:
                MoveLeft := TRUE;
                actionInProgress := TRUE;
                IF LeftLimitSwitch THEN
                    MoveLeft := FALSE;
                    actionInProgress := FALSE;
                    stepNumber := 1;
                END_IF;
        END_CASE;
    END_IF;
END_IF;
END_FUNCTION_BLOCK
